      W_g[13,37] := -0.07636662;
      W_g[13,38] := -0.02541909;
      W_g[13,39] := -0.00815807;
      W_g[14,0] := 0.05384851;
      W_g[14,1] := -0.08540776;
      W_g[14,2] := -0.08017597;
      W_g[14,3] := -0.28711280;
      W_g[14,4] := -0.38180253;
      W_g[14,5] := -0.12807073;
      W_g[14,6] := -0.33112118;
      W_g[14,7] := -0.01536665;
      W_g[14,8] := 0.07860034;
      W_g[14,9] := 0.07597807;
      W_g[14,10] := 0.81271881;
      W_g[14,11] := 0.34440023;
      W_g[14,12] := -0.11264267;
      W_g[14,13] := 0.29767352;
      W_g[14,14] := -0.05823113;
      W_g[14,15] := -0.00107844;
      W_g[14,16] := -0.02762355;
      W_g[14,17] := -0.02232336;
      W_g[14,18] := 0.03123496;
      W_g[14,19] := -0.13857344;
      W_g[14,20] := 0.10911304;
      W_g[14,21] := -0.12785229;
      W_g[14,22] := -0.04815350;
      W_g[14,23] := -0.17390981;
      W_g[14,24] := 0.13923632;
      W_g[14,25] := 0.11850380;
      W_g[14,26] := -0.32757759;
      W_g[14,27] := -0.25137767;
      W_g[14,28] := 0.22421645;
      W_g[14,29] := -0.42832899;
      W_g[14,30] := 0.06481594;
      W_g[14,31] := -0.23915793;
      W_g[14,32] := -0.04046796;
      W_g[14,33] := -0.09582479;
      W_g[14,34] := -0.09370243;
      W_g[14,35] := 0.14524275;
      W_g[14,36] := -0.03895468;
      W_g[14,37] := 0.10286443;
      W_g[14,38] := 0.03800159;
      W_g[14,39] := 0.11008195;
      W_g[15,0] := 0.49670509;
      W_g[15,1] := 0.19451231;
      W_g[15,2] := -0.24881296;
      W_g[15,3] := 0.56299460;
      W_g[15,4] := -0.14983681;
      W_g[15,5] := -0.02904006;
      W_g[15,6] := 0.06259420;
      W_g[15,7] := 0.16642898;
      W_g[15,8] := -0.08521152;
      W_g[15,9] := -0.12409624;
      W_g[15,10] := 0.24281517;
      W_g[15,11] := -0.10940242;
      W_g[15,12] := 0.71269953;
      W_g[15,13] := -0.18780579;
      W_g[15,14] := 0.00091037;
      W_g[15,15] := -0.06534981;
      W_g[15,16] := 0.00326133;
      W_g[15,17] := -0.00118504;
      W_g[15,18] := -0.04420842;
      W_g[15,19] := -0.22520956;
      W_g[15,20] := -0.11959776;
      W_g[15,21] := -0.10079119;
      W_g[15,22] := -0.04329386;
      W_g[15,23] := -0.07395163;
      W_g[15,24] := -0.11715485;
      W_g[15,25] := -0.18832952;
      W_g[15,26] := -0.24700920;
      W_g[15,27] := -0.09096922;
      W_g[15,28] := 0.07692285;
      W_g[15,29] := 0.01714239;
      W_g[15,30] := -0.08180999;
      W_g[15,31] := -0.00006038;
      W_g[15,32] := 0.02792178;
      W_g[15,33] := 0.08978129;
      W_g[15,34] := -0.02846152;
      W_g[15,35] := 0.05397168;
      W_g[15,36] := 0.01382420;
      W_g[15,37] := 0.12623927;
      W_g[15,38] := 0.02842882;
      W_g[15,39] := -0.23873122;
      W_g[16,0] := 0.00714069;
      W_g[16,1] := 0.09252225;
      W_g[16,2] := -0.01911032;
      W_g[16,3] := 0.04820935;
      W_g[16,4] := 0.04210250;
      W_g[16,5] := 0.05442985;
      W_g[16,6] := 0.24199863;
      W_g[16,7] := -0.08810946;
      W_g[16,8] := 0.02272573;
      W_g[16,9] := -0.01153773;
      W_g[16,10] := -0.01938002;
      W_g[16,11] := 0.95534259;
      W_g[16,12] := 0.00685452;
      W_g[16,13] := -0.05267539;
      W_g[16,14] := -0.04784015;
      W_g[16,15] := 0.02123881;
      W_g[16,16] := 0.02990256;
      W_g[16,17] := 0.22012618;
      W_g[16,18] := -0.12446024;
      W_g[16,19] := 0.01318580;
      W_g[16,20] := 0.31736228;
      W_g[16,21] := 0.25552613;
      W_g[16,22] := 0.02996899;
      W_g[16,23] := 0.13324806;
      W_g[16,24] := 0.01029211;
      W_g[16,25] := -0.11731086;
      W_g[16,26] := 0.08171849;
      W_g[16,27] := -0.11919475;
      W_g[16,28] := 0.04512075;
      W_g[16,29] := 0.04511562;
      W_g[16,30] := 0.01768237;
      W_g[16,31] := -0.11807074;
      W_g[16,32] := 0.02917237;
      W_g[16,33] := 0.08451862;
      W_g[16,34] := 0.18420373;
      W_g[16,35] := 0.06097095;
      W_g[16,36] := 0.01656622;
      W_g[16,37] := -0.02950481;
      W_g[16,38] := 0.00875620;
      W_g[16,39] := -0.30139515;
      W_g[17,0] := 0.28211352;
      W_g[17,1] := -0.06947739;
      W_g[17,2] := -0.48255709;
      W_g[17,3] := -0.48009890;
      W_g[17,4] := 0.40037093;
      W_g[17,5] := -0.41533524;
      W_g[17,6] := 0.61539871;
      W_g[17,7] := -0.07803038;
      W_g[17,8] := 0.20740844;
      W_g[17,9] := 0.19454060;
      W_g[17,10] := 0.37828967;
      W_g[17,11] := 0.51134646;
      W_g[17,12] := 0.02942824;
      W_g[17,13] := -0.03419436;
      W_g[17,14] := -0.14622004;
      W_g[17,15] := 0.12808461;
      W_g[17,16] := -0.08771772;
      W_g[17,17] := -0.17915098;
      W_g[17,18] := -0.35652786;
      W_g[17,19] := -0.08436973;
      W_g[17,20] := -0.15241621;
      W_g[17,21] := -0.59241575;
      W_g[17,22] := -0.12622987;
      W_g[17,23] := -0.06875754;
      W_g[17,24] := -0.61650282;
      W_g[17,25] := -0.62400168;
      W_g[17,26] := 0.12978441;
      W_g[17,27] := 0.19093341;
      W_g[17,28] := -0.57437402;
      W_g[17,29] := -0.10343723;
      W_g[17,30] := -0.14047481;
      W_g[17,31] := 0.10861561;
      W_g[17,32] := -0.08338292;
      W_g[17,33] := -0.15795745;
      W_g[17,34] := -1.05674601;
      W_g[17,35] := 0.07798125;
      W_g[17,36] := -0.04106956;
      W_g[17,37] := -0.14353254;
      W_g[17,38] := -0.01768998;
      W_g[17,39] := 0.23552968;
      W_g[18,0] := -0.56118143;
      W_g[18,1] := 0.01680752;
      W_g[18,2] := 0.21060835;
      W_g[18,3] := 0.22311090;
      W_g[18,4] := -0.35391527;
      W_g[18,5] := -0.00398842;
      W_g[18,6] := 0.44133097;
      W_g[18,7] := -0.20236395;
      W_g[18,8] := 0.27059153;
      W_g[18,9] := -0.26535335;
      W_g[18,10] := -0.00161409;
      W_g[18,11] := -0.42498562;
      W_g[18,12] := 0.18595842;
      W_g[18,13] := 0.03403796;
      W_g[18,14] := -0.19036941;
      W_g[18,15] := 0.00153053;
      W_g[18,16] := -0.13208415;
      W_g[18,17] := -0.00688618;
      W_g[18,18] := 0.04695740;
      W_g[18,19] := 0.52580279;
      W_g[18,20] := 0.33302781;
      W_g[18,21] := -0.03863472;
      W_g[18,22] := -0.04098545;
      W_g[18,23] := 0.05270698;
      W_g[18,24] := -0.87936115;
      W_g[18,25] := -0.79176319;
      W_g[18,26] := -0.37981445;
      W_g[18,27] := -0.39054155;
      W_g[18,28] := 0.40099201;
      W_g[18,29] := -0.21964216;
      W_g[18,30] := -0.06956752;
      W_g[18,31] := 1.08965826;
      W_g[18,32] := -0.24863915;
      W_g[18,33] := 0.04124767;
      W_g[18,34] := -0.14617871;
      W_g[18,35] := -0.54955792;
      W_g[18,36] := 0.22360204;
      W_g[18,37] := -0.51476938;
      W_g[18,38] := -0.00649375;
      W_g[18,39] := 0.23745580;
      W_g[19,0] := 0.04427215;
      W_g[19,1] := 0.13209015;
      W_g[19,2] := -0.12966105;
      W_g[19,3] := 0.13671713;
      W_g[19,4] := 0.01762369;
      W_g[19,5] := 0.09627694;
      W_g[19,6] := -0.13640797;
      W_g[19,7] := 0.02292525;
      W_g[19,8] := 0.06818993;
      W_g[19,9] := -0.01616117;
      W_g[19,10] := -0.27115190;
      W_g[19,11] := -0.17511748;
      W_g[19,12] := 0.20083658;
      W_g[19,13] := 0.12117302;
      W_g[19,14] := -0.40477425;
      W_g[19,15] := 0.00942509;
      W_g[19,16] := -0.00977145;
      W_g[19,17] := -0.00656325;
      W_g[19,18] := -0.02440832;
      W_g[19,19] := -0.10208004;
      W_g[19,20] := 0.05442004;
      W_g[19,21] := -0.28210428;
      W_g[19,22] := -0.02802154;
      W_g[19,23] := -0.16558743;
      W_g[19,24] := 0.24839798;
      W_g[19,25] := 0.68076271;
      W_g[19,26] := -0.15649894;
      W_g[19,27] := 0.02872765;
      W_g[19,28] := -0.14855081;
      W_g[19,29] := -0.04783039;
      W_g[19,30] := -0.04433315;
      W_g[19,31] := -0.00463518;
      W_g[19,32] := -0.04792630;
      W_g[19,33] := -0.18936750;
      W_g[19,34] := -0.28109401;
      W_g[19,35] := 0.12269117;
      W_g[19,36] := -0.02590044;
      W_g[19,37] := 0.13191973;
      W_g[19,38] := -0.08906776;
      W_g[19,39] := -0.30020091;
      W_g[20,0] := -0.20718005;
      W_g[20,1] := -0.84034145;
      W_g[20,2] := 0.02167286;
      W_g[20,3] := 0.22337365;
      W_g[20,4] := -0.22535181;
      W_g[20,5] := 0.00862414;
      W_g[20,6] := -0.07585888;
      W_g[20,7] := 0.20224823;
      W_g[20,8] := 0.33609936;
      W_g[20,9] := 0.24086921;
      W_g[20,10] := -0.34230143;
      W_g[20,11] := 0.23271726;
      W_g[20,12] := -0.54696190;
      W_g[20,13] := 0.07557353;
      W_g[20,14] := -0.00750887;
      W_g[20,15] := -0.07179558;
      W_g[20,16] := 0.11929045;
      W_g[20,17] := 0.01187360;
      W_g[20,18] := 0.01727761;
      W_g[20,19] := -0.10120918;
      W_g[20,20] := -0.35278231;
      W_g[20,21] := -0.09405834;
      W_g[20,22] := 0.04689666;
      W_g[20,23] := -0.10715894;
      W_g[20,24] := -0.07375087;
      W_g[20,25] := -0.14543816;
      W_g[20,26] := -0.23896208;
      W_g[20,27] := -0.43519315;
      W_g[20,28] := -0.25828305;
      W_g[20,29] := -0.05447736;
      W_g[20,30] := 0.05642707;
      W_g[20,31] := 0.18183576;
      W_g[20,32] := 0.08492490;
      W_g[20,33] := 0.19067700;
      W_g[20,34] := -0.11871803;
      W_g[20,35] := -0.03175204;
      W_g[20,36] := -0.04638923;
      W_g[20,37] := -0.03955484;
      W_g[20,38] := 0.18262649;
      W_g[20,39] := -0.00053967;
      W_g[21,0] := -0.00852127;
      W_g[21,1] := 0.16749823;
      W_g[21,2] := -0.15172872;
      W_g[21,3] := -0.20800257;
      W_g[21,4] := 0.15032937;
      W_g[21,5] := 0.06710505;
      W_g[21,6] := -0.26149949;
      W_g[21,7] := 0.03740874;
      W_g[21,8] := 0.13018388;
      W_g[21,9] := 0.18329854;
      W_g[21,10] := -0.03891287;
      W_g[21,11] := 0.05188271;
      W_g[21,12] := 0.47803098;
      W_g[21,13] := 0.06662370;
      W_g[21,14] := -0.00612103;
      W_g[21,15] := -0.13870122;
      W_g[21,16] := -0.10494442;
      W_g[21,17] := -0.00346555;
      W_g[21,18] := -0.04227602;
      W_g[21,19] := -0.33476129;
      W_g[21,20] := 0.34089175;
      W_g[21,21] := 0.45425063;
      W_g[21,22] := 0.16435136;
      W_g[21,23] := 0.04143468;
      W_g[21,24] := 0.16786721;
      W_g[21,25] := 0.11948983;
      W_g[21,26] := 0.05792047;
      W_g[21,27] := -0.12976640;
      W_g[21,28] := -0.13790442;
      W_g[21,29] := 0.24387960;
      W_g[21,30] := 0.16521277;
      W_g[21,31] := 0.16834626;
      W_g[21,32] := -0.10805231;
      W_g[21,33] := -0.07898282;
      W_g[21,34] := 0.28881353;
      W_g[21,35] := -0.11385613;
      W_g[21,36] := -0.66726488;
      W_g[21,37] := -0.28654984;
      W_g[21,38] := 0.35271052;
      W_g[21,39] := 0.00955431;
      W_g[22,0] := 0.29109696;
      W_g[22,1] := 0.01384218;
      W_g[22,2] := -0.37709463;
      W_g[22,3] := 0.14574254;
      W_g[22,4] := -0.07661973;
      W_g[22,5] := 0.12081382;
      W_g[22,6] := -0.39220569;
      W_g[22,7] := -0.00977318;
      W_g[22,8] := 0.02812388;
      W_g[22,9] := -0.07591717;
      W_g[22,10] := -0.08413436;
      W_g[22,11] := 0.17591499;
      W_g[22,12] := -0.33312052;
      W_g[22,13] := -0.12893844;
      W_g[22,14] := 0.12280960;
      W_g[22,15] := 0.33149692;
      W_g[22,16] := -0.12770943;
      W_g[22,17] := 0.11019890;
      W_g[22,18] := -0.02004679;
      W_g[22,19] := -0.09840271;
      W_g[22,20] := -0.03289499;
      W_g[22,21] := -0.03317460;
      W_g[22,22] := 0.05239879;
      W_g[22,23] := 0.39912307;
      W_g[22,24] := 0.28896907;
      W_g[22,25] := -0.06105658;
      W_g[22,26] := -0.21285506;
      W_g[22,27] := -0.03863349;
      W_g[22,28] := 0.16256362;
      W_g[22,29] := 0.14152323;
      W_g[22,30] := 0.05700575;
      W_g[22,31] := 0.37323594;
      W_g[22,32] := -0.00197801;
      W_g[22,33] := 0.01016807;
      W_g[22,34] := -0.05393393;
      W_g[22,35] := -0.03373878;
      W_g[22,36] := 0.00123443;
      W_g[22,37] := -0.10641941;
      W_g[22,38] := -0.03629038;
      W_g[22,39] := -0.09397990;
      W_g[23,0] := -0.09347695;
      W_g[23,1] := -0.22505829;
      W_g[23,2] := 0.01111710;
      W_g[23,3] := -0.13649231;
      W_g[23,4] := -0.30517000;
      W_g[23,5] := 0.83911264;
      W_g[23,6] := -0.75282311;
      W_g[23,7] := -0.66691148;
      W_g[23,8] := 0.15447931;
      W_g[23,9] := -0.55708647;
      W_g[23,10] := 0.25686628;
      W_g[23,11] := 0.12212675;
      W_g[23,12] := 0.16343321;
      W_g[23,13] := -0.31660068;
      W_g[23,14] := 0.02282131;
      W_g[23,15] := -0.05205119;
      W_g[23,16] := -0.05839873;
      W_g[23,17] := -0.09075660;
      W_g[23,18] := -0.23147778;
      W_g[23,19] := 0.07263616;
      W_g[23,20] := -0.51794368;
      W_g[23,21] := -0.27791360;
      W_g[23,22] := -0.07805633;
      W_g[23,23] := -0.41355452;
      W_g[23,24] := -0.21751262;
      W_g[23,25] := -0.05684796;
      W_g[23,26] := 0.30686048;
      W_g[23,27] := -0.14003992;
      W_g[23,28] := -0.38135511;
      W_g[23,29] := 0.13330600;
      W_g[23,30] := -0.06790695;
      W_g[23,31] := -0.07987443;
      W_g[23,32] := 0.06365003;
      W_g[23,33] := 0.22799088;
      W_g[23,34] := 0.13270302;
      W_g[23,35] := -0.00725970;
      W_g[23,36] := 0.16376778;
      W_g[23,37] := -0.02287991;
      W_g[23,38] := 0.08711061;
      W_g[23,39] := 0.01950686;
      W_g[24,0] := 0.46194655;
      W_g[24,1] := 0.27763960;
      W_g[24,2] := -0.12869456;
      W_g[24,3] := 0.13782990;
      W_g[24,4] := -1.03041399;
      W_g[24,5] := 0.00441816;
      W_g[24,6] := 0.44230226;
      W_g[24,7] := 0.18489341;
      W_g[24,8] := -0.30371043;
      W_g[24,9] := 0.03693367;
      W_g[24,10] := -0.01524317;
      W_g[24,11] := -0.24215870;
      W_g[24,12] := 0.35080424;
      W_g[24,13] := 0.07174128;
      W_g[24,14] := 0.00412538;
      W_g[24,15] := 0.02062515;
      W_g[24,16] := 0.01971583;
      W_g[24,17] := 0.00580471;
      W_g[24,18] := -0.04475251;
      W_g[24,19] := -0.08863095;
      W_g[24,20] := 0.06659620;
      W_g[24,21] := -0.19372395;
      W_g[24,22] := 0.04916465;
      W_g[24,23] := 0.11263776;
      W_g[24,24] := 0.45533353;
      W_g[24,25] := 0.28435835;
      W_g[24,26] := 0.23480317;
      W_g[24,27] := -0.41078931;
      W_g[24,28] := -0.25990930;
      W_g[24,29] := 0.04082377;
      W_g[24,30] := 0.05907518;
      W_g[24,31] := 0.00033808;
      W_g[24,32] := -0.03658906;
      W_g[24,33] := -0.08924066;
      W_g[24,34] := -0.02038150;
      W_g[24,35] := 0.01517213;
      W_g[24,36] := -0.29084125;
      W_g[24,37] := -0.03483975;
      W_g[24,38] := -0.33877048;
      W_g[24,39] := 0.01846378;
      W_g[25,0] := -0.01319884;
      W_g[25,1] := 0.17892542;
      W_g[25,2] := 0.00354903;
      W_g[25,3] := -0.01092031;
      W_g[25,4] := 0.04581180;
      W_g[25,5] := -0.04252854;
      W_g[25,6] := -0.05655812;
      W_g[25,7] := 0.07682356;
      W_g[25,8] := -0.01679150;
      W_g[25,9] := 0.05484685;
      W_g[25,10] := -0.09173104;
      W_g[25,11] := -0.12738757;
      W_g[25,12] := -0.10293069;
      W_g[25,13] := -0.00530847;
      W_g[25,14] := -0.08904938;
      W_g[25,15] := 0.36966512;
      W_g[25,16] := -0.00969987;
      W_g[25,17] := -0.28969538;
      W_g[25,18] := -0.02469883;
      W_g[25,19] := -0.08574332;
      W_g[25,20] := 0.10813141;
      W_g[25,21] := 0.08889347;
      W_g[25,22] := -0.06467538;
      W_g[25,23] := 0.04102366;
      W_g[25,24] := -0.24661052;
      W_g[25,25] := -0.24702097;
      W_g[25,26] := -0.08217103;
      W_g[25,27] := -0.05707087;
      W_g[25,28] := -0.01940200;
      W_g[25,29] := -0.00729063;
      W_g[25,30] := -0.06900500;
      W_g[25,31] := -0.19478676;
      W_g[25,32] := 0.08665588;
      W_g[25,33] := 0.17711434;
      W_g[25,34] := 0.35117847;
      W_g[25,35] := 0.00400291;
      W_g[25,36] := 0.02780187;
      W_g[25,37] := -0.02507502;
      W_g[25,38] := 0.01814217;
      W_g[25,39] := 0.01270028;
      W_g[26,0] := -0.10013371;
      W_g[26,1] := -0.11928739;
      W_g[26,2] := 0.03542966;
      W_g[26,3] := -0.09299100;
      W_g[26,4] := 0.22154348;
      W_g[26,5] := 0.04870279;
      W_g[26,6] := -0.01336484;
      W_g[26,7] := -0.05781888;
      W_g[26,8] := 0.00065369;
      W_g[26,9] := -0.01473211;
      W_g[26,10] := -0.01971318;
      W_g[26,11] := 0.02451181;
      W_g[26,12] := 0.14100704;
      W_g[26,13] := 0.20081082;
      W_g[26,14] := -0.00175938;
      W_g[26,15] := -0.13420245;
      W_g[26,16] := 0.01900839;
      W_g[26,17] := -0.02341681;
      W_g[26,18] := -0.94101948;
      W_g[26,19] := -0.02586854;
      W_g[26,20] := -0.30304915;
      W_g[26,21] := 0.06037450;
      W_g[26,22] := -0.02225667;
      W_g[26,23] := 0.34992269;
      W_g[26,24] := -0.15178578;
      W_g[26,25] := -0.21104257;
      W_g[26,26] := -0.25511426;
      W_g[26,27] := -0.03610617;
      W_g[26,28] := -0.13982570;
      W_g[26,29] := -0.07677662;
      W_g[26,30] := -0.02899644;
      W_g[26,31] := 0.02322534;
      W_g[26,32] := -0.01148466;
      W_g[26,33] := 0.01643471;
      W_g[26,34] := -0.05193237;
      W_g[26,35] := -0.01343275;
      W_g[26,36] := 0.01284295;
      W_g[26,37] := 0.01176736;
      W_g[26,38] := 0.00468252;
      W_g[26,39] := -0.20358260;
      W_g[27,0] := 0.01242287;
      W_g[27,1] := -0.01930982;
      W_g[27,2] := -0.24737412;
      W_g[27,3] := -0.13776387;
      W_g[27,4] := 0.19126348;
      W_g[27,5] := 0.00086061;
      W_g[27,6] := -0.16852112;
      W_g[27,7] := -0.08134060;
      W_g[27,8] := 0.29883468;
      W_g[27,9] := 0.09754812;
      W_g[27,10] := 0.09034698;
      W_g[27,11] := -0.06812658;
      W_g[27,12] := -0.14695419;
      W_g[27,13] := -0.05109974;
      W_g[27,14] := -0.01788860;
      W_g[27,15] := -0.15783192;
      W_g[27,16] := 0.19530444;
      W_g[27,17] := -0.16005373;
      W_g[27,18] := 0.26013258;
      W_g[27,19] := 0.26764771;
      W_g[27,20] := -0.12696983;
      W_g[27,21] := 0.31249490;
      W_g[27,22] := 0.09300645;
      W_g[27,23] := 0.03466551;
      W_g[27,24] := 0.23168693;
      W_g[27,25] := 0.18956751;
      W_g[27,26] := -0.04334988;
      W_g[27,27] := -0.18214862;
      W_g[27,28] := -0.04629618;
      W_g[27,29] := 0.09379144;
      W_g[27,30] := 0.07671305;
      W_g[27,31] := -0.01221954;
      W_g[27,32] := -0.02424719;
      W_g[27,33] := 0.07423434;
      W_g[27,34] := 0.18019708;
      W_g[27,35] := -0.04701952;
      W_g[27,36] := -0.08283819;
      W_g[27,37] := -0.09333491;
      W_g[27,38] := -0.48927879;
      W_g[27,39] := -0.00745687;
      W_g[28,0] := 0.13821959;
      W_g[28,1] := 0.07419970;
      W_g[28,2] := -0.28731343;
      W_g[28,3] := 0.52230597;
      W_g[28,4] := 0.13792820;
      W_g[28,5] := -0.04003582;
      W_g[28,6] := 0.12009837;
      W_g[28,7] := -0.22427090;
      W_g[28,8] := 0.10034105;
      W_g[28,9] := -0.43725863;
      W_g[28,10] := 0.10780185;
      W_g[28,11] := -0.03007025;
      W_g[28,12] := -0.09082274;
      W_g[28,13] := 0.21732096;
      W_g[28,14] := -0.03366475;
      W_g[28,15] := 0.12757394;
      W_g[28,16] := 0.40819040;
      W_g[28,17] := 0.08709385;
      W_g[28,18] := -0.01960146;
      W_g[28,19] := -0.01771599;
      W_g[28,20] := 0.02389354;
      W_g[28,21] := 0.04893105;
      W_g[28,22] := 0.01708278;
      W_g[28,23] := 0.05532730;
      W_g[28,24] := -0.42513239;
      W_g[28,25] := -0.53693467;
      W_g[28,26] := 0.09680068;
      W_g[28,27] := 0.11012019;
      W_g[28,28] := -0.10853667;
      W_g[28,29] := -0.10696560;
      W_g[28,30] := -0.01152095;
      W_g[28,31] := 0.08765919;
      W_g[28,32] := -0.04124034;
      W_g[28,33] := 0.00073121;
      W_g[28,34] := -0.07680846;
      W_g[28,35] := -0.09583755;
      W_g[28,36] := -0.02250235;
      W_g[28,37] := -0.10466012;
      W_g[28,38] := 0.02804276;
      W_g[28,39] := 0.05010757;
      W_g[29,0] := -0.13576494;
      W_g[29,1] := -0.04743524;
      W_g[29,2] := 0.01165335;
      W_g[29,3] := -0.06858198;
      W_g[29,4] := 0.11698179;
      W_g[29,5] := 0.15293106;
      W_g[29,6] := -0.08868138;
      W_g[29,7] := 0.00604072;
      W_g[29,8] := 0.10700601;
      W_g[29,9] := 0.08990686;
      W_g[29,10] := -0.17016383;
      W_g[29,11] := -0.09298281;
      W_g[29,12] := 0.23396063;
      W_g[29,13] := -0.43684760;
      W_g[29,14] := -0.02256006;
      W_g[29,15] := 0.02156748;
      W_g[29,16] := -0.04530424;
      W_g[29,17] := 0.02112582;
      W_g[29,18] := 0.43311554;
      W_g[29,19] := 0.28956264;
      W_g[29,20] := -0.45648861;
      W_g[29,21] := -0.47465628;
      W_g[29,22] := -0.15953651;
      W_g[29,23] := 0.62224460;
      W_g[29,24] := -0.36037850;
      W_g[29,25] := -0.32347810;
      W_g[29,26] := -0.10036322;
      W_g[29,27] := 0.23475674;
      W_g[29,28] := -0.38871291;
      W_g[29,29] := -0.37588716;
      W_g[29,30] := -0.19999301;
      W_g[29,31] := -0.07129297;
      W_g[29,32] := 0.00924866;
      W_g[29,33] := -0.00100953;
      W_g[29,34] := -0.03974389;
      W_g[29,35] := 0.19243315;
      W_g[29,36] := -0.05763126;
      W_g[29,37] := 0.14980933;
      W_g[29,38] := 0.09773512;
      W_g[29,39] := 0.28358760;
      W_g[30,0] := 0.02073097;
      W_g[30,1] := -0.05142897;
      W_g[30,2] := 0.05679109;
      W_g[30,3] := -0.29680440;
      W_g[30,4] := -0.09398746;
      W_g[30,5] := 0.00418108;
      W_g[30,6] := -0.12116858;
      W_g[30,7] := 0.13785014;
      W_g[30,8] := -0.07182530;
      W_g[30,9] := 0.28989494;
      W_g[30,10] := -0.02703100;
      W_g[30,11] := -0.04196686;
      W_g[30,12] := 0.23686379;
      W_g[30,13] := -0.11817347;
      W_g[30,14] := -0.00608444;
      W_g[30,15] := 0.27866739;
      W_g[30,16] := 0.31624600;
      W_g[30,17] := -0.04371030;
      W_g[30,18] := -0.09872175;
      W_g[30,19] := 0.17183733;
      W_g[30,20] := -0.10328431;
      W_g[30,21] := 0.02654029;
      W_g[30,22] := 0.04664133;
      W_g[30,23] := -0.02138521;
      W_g[30,24] := 0.42544174;
      W_g[30,25] := -0.03961691;
      W_g[30,26] := 0.11087703;
      W_g[30,27] := 0.09755427;
      W_g[30,28] := 0.11475538;
      W_g[30,29] := 0.06603787;
      W_g[30,30] := 0.05809331;
      W_g[30,31] := 0.13511968;
      W_g[30,32] := -0.00735715;
      W_g[30,33] := -0.00152808;
      W_g[30,34] := -0.12982640;
      W_g[30,35] := 0.00118882;
      W_g[30,36] := 0.01855830;
      W_g[30,37] := -0.05438844;
      W_g[30,38] := 0.05046400;
      W_g[30,39] := -0.03010074;
      W_g[31,0] := 0.08256169;
      W_g[31,1] := -0.51133311;
      W_g[31,2] := 0.11336197;
      W_g[31,3] := -0.15730928;
      W_g[31,4] := 0.15212694;
      W_g[31,5] := 0.05411269;
      W_g[31,6] := -0.07535803;
      W_g[31,7] := 0.03512096;
      W_g[31,8] := -0.05313810;
      W_g[31,9] := 0.10365095;
      W_g[31,10] := -0.00368842;
      W_g[31,11] := -0.12890872;
      W_g[31,12] := 0.47981134;
      W_g[31,13] := 0.03815160;
      W_g[31,14] := -0.01872904;
      W_g[31,15] := 0.17062889;
      W_g[31,16] := -0.12828785;
      W_g[31,17] := 0.06558654;
      W_g[31,18] := -0.06244295;
      W_g[31,19] := -0.53075397;
      W_g[31,20] := 0.15929437;
      W_g[31,21] := 0.00589449;
      W_g[31,22] := -0.03731958;
      W_g[31,23] := 0.05464490;
      W_g[31,24] := -0.19547676;
      W_g[31,25] := 0.11578897;
      W_g[31,26] := 0.27690557;
      W_g[31,27] := 0.26996168;
      W_g[31,28] := 0.03783383;
      W_g[31,29] := -0.16668507;
      W_g[31,30] := -0.05871727;
      W_g[31,31] := 0.11560699;
      W_g[31,32] := -0.10597849;
      W_g[31,33] := -0.03747635;
      W_g[31,34] := -0.06264409;
      W_g[31,35] := -0.18381201;
      W_g[31,36] := 0.07526756;
      W_g[31,37] := -0.11970815;
      W_g[31,38] := -0.33985323;
      W_g[31,39] := 0.02983656;
      W_o[0,0] := 0.13366428;
      W_o[0,1] := 0.11036980;
      W_o[0,2] := -0.16846675;
      W_o[0,3] := -0.21495235;
      W_o[0,4] := 0.07811608;
      W_o[0,5] := -0.13181226;
      W_o[0,6] := -0.32309711;
      W_o[0,7] := -0.05775660;
      W_o[0,8] := 0.07714970;
      W_o[0,9] := 0.69965583;
      W_o[0,10] := 0.03330577;
      W_o[0,11] := 0.07725812;
      W_o[0,12] := 0.25551820;
      W_o[0,13] := 0.38036522;
      W_o[0,14] := -0.01993838;
      W_o[0,15] := -0.05171372;
      W_o[0,16] := 0.00189644;
      W_o[0,17] := -0.32097366;
      W_o[0,18] := -0.05273939;
      W_o[0,19] := 0.04321737;
      W_o[0,20] := -0.23801146;
      W_o[0,21] := 0.29699677;
      W_o[0,22] := -0.16276316;
      W_o[0,23] := -0.23706993;
      W_o[0,24] := 0.17703076;
      W_o[0,25] := 0.36713782;
      W_o[0,26] := -0.12915254;
      W_o[0,27] := -0.07524700;
      W_o[0,28] := -0.09860305;
      W_o[0,29] := 0.12421684;
      W_o[0,30] := -0.39039981;
      W_o[0,31] := -0.01002511;
      W_o[0,32] := -0.46100792;
      W_o[0,33] := 0.17252544;
      W_o[0,34] := 0.15642625;
      W_o[0,35] := -0.27402765;
      W_o[0,36] := -0.07788435;
      W_o[0,37] := -0.09713101;
      W_o[0,38] := -0.05069508;
      W_o[0,39] := -0.24549620;
      W_o[1,0] := 0.49653649;
      W_o[1,1] := -0.05346184;
      W_o[1,2] := -0.01993282;
      W_o[1,3] := -0.13199322;
      W_o[1,4] := 0.03771848;
      W_o[1,5] := 0.14309798;
      W_o[1,6] := 0.04961836;
      W_o[1,7] := 0.27153552;
      W_o[1,8] := 0.60058177;
      W_o[1,9] := -0.62969673;
      W_o[1,10] := 0.21819758;
      W_o[1,11] := -0.10272143;
      W_o[1,12] := 0.11986823;
      W_o[1,13] := -0.24452005;
      W_o[1,14] := -0.06335072;
      W_o[1,15] := -0.16848719;
      W_o[1,16] := -0.21195354;
      W_o[1,17] := 0.02550812;
      W_o[1,18] := -0.14588526;
      W_o[1,19] := -0.51397264;
      W_o[1,20] := -0.21644965;
      W_o[1,21] := -0.53661948;
      W_o[1,22] := -0.02092957;
      W_o[1,23] := 0.01972848;
      W_o[1,24] := -0.55939800;
      W_o[1,25] := -0.49083781;
      W_o[1,26] := -0.14633974;
      W_o[1,27] := 0.42070836;
      W_o[1,28] := -0.21612938;
      W_o[1,29] := -0.03745779;
      W_o[1,30] := 0.06127948;
      W_o[1,31] := 0.35676870;
      W_o[1,32] := -0.08789702;
      W_o[1,33] := 0.11810053;
      W_o[1,34] := -0.01725286;
      W_o[1,35] := -0.06969324;
      W_o[1,36] := -0.01398361;
      W_o[1,37] := -0.15410708;
      W_o[1,38] := -0.08071988;
      W_o[1,39] := -0.25934911;
      W_o[2,0] := 0.13397244;
      W_o[2,1] := -0.67044854;
      W_o[2,2] := -0.32567781;
      W_o[2,3] := -0.75043666;
      W_o[2,4] := -0.32291642;
      W_o[2,5] := 0.54297352;
      W_o[2,6] := 1.01406825;
      W_o[2,7] := -0.63293743;
      W_o[2,8] := -0.24675053;
      W_o[2,9] := -0.54400074;
      W_o[2,10] := -0.70754099;
      W_o[2,11] := -0.16770625;
      W_o[2,12] := -0.13771380;
      W_o[2,13] := -0.93835974;
      W_o[2,14] := 0.07016375;
      W_o[2,15] := -0.14486392;
      W_o[2,16] := 0.26753914;
      W_o[2,17] := -0.44003579;
      W_o[2,18] := -0.19662693;
      W_o[2,19] := 0.14748774;
      W_o[2,20] := 0.04340832;
      W_o[2,21] := 0.91405821;
      W_o[2,22] := 0.23963371;
      W_o[2,23] := -0.42069820;
      W_o[2,24] := 1.35907292;
      W_o[2,25] := 0.74127895;
      W_o[2,26] := -0.60126311;
      W_o[2,27] := 1.04573679;
      W_o[2,28] := 0.35571697;
      W_o[2,29] := 0.19770171;
      W_o[2,30] := 0.19496830;
      W_o[2,31] := -0.06545950;
      W_o[2,32] := -0.07142299;
      W_o[2,33] := -0.23412317;
      W_o[2,34] := 0.13213682;
      W_o[2,35] := 0.09960951;
      W_o[2,36] := -0.82927501;
      W_o[2,37] := -0.00553483;
      W_o[2,38] := 0.72544241;
      W_o[2,39] := 0.20440662;
      W_o[3,0] := -0.29025504;
      W_o[3,1] := 0.21485890;
      W_o[3,2] := 0.12162556;
      W_o[3,3] := -0.45000923;
      W_o[3,4] := 0.00440878;
      W_o[3,5] := -0.07761150;
      W_o[3,6] := 0.27128229;
      W_o[3,7] := 0.20583764;
      W_o[3,8] := 0.36606720;
      W_o[3,9] := 0.31630817;
      W_o[3,10] := 0.16728929;
      W_o[3,11] := 0.21024089;
      W_o[3,12] := -0.30256730;
      W_o[3,13] := -0.07960982;
      W_o[3,14] := 0.26832253;
      W_o[3,15] := 0.38332802;
      W_o[3,16] := 0.01548071;
      W_o[3,17] := 0.27411333;
      W_o[3,18] := -0.07721005;
      W_o[3,19] := -0.15753639;
      W_o[3,20] := -0.12283424;
      W_o[3,21] := -0.09994975;
      W_o[3,22] := -0.25781667;
      W_o[3,23] := -0.30848202;
      W_o[3,24] := 0.08977263;
      W_o[3,25] := -0.00644524;
      W_o[3,26] := 0.31200859;
      W_o[3,27] := -0.01467965;
      W_o[3,28] := -0.12804723;
      W_o[3,29] := -0.06573117;
      W_o[3,30] := -0.39431822;
      W_o[3,31] := -0.44901580;
      W_o[3,32] := -0.13384379;
      W_o[3,33] := -0.10575464;
      W_o[3,34] := 0.01442572;
      W_o[3,35] := -0.11673454;
      W_o[3,36] := -0.14822102;
      W_o[3,37] := -0.02524356;
      W_o[3,38] := -0.03832110;
      W_o[3,39] := 0.94678485;
      W_o[4,0] := -0.89165902;
      W_o[4,1] := -0.07221486;
      W_o[4,2] := 0.45090771;
      W_o[4,3] := 0.40743887;
      W_o[4,4] := -0.00022854;
      W_o[4,5] := -0.22787750;
      W_o[4,6] := 0.56126112;
      W_o[4,7] := -0.65236539;
      W_o[4,8] := 0.31672934;
      W_o[4,9] := -0.60582823;
      W_o[4,10] := 0.85605830;
      W_o[4,11] := -0.86477047;
      W_o[4,12] := 0.63425988;
      W_o[4,13] := -0.08753718;
      W_o[4,14] := 0.07426148;
      W_o[4,15] := 0.43497530;
      W_o[4,16] := 0.02985676;
      W_o[4,17] := -0.01102423;
      W_o[4,18] := 0.00179447;
      W_o[4,19] := -0.39584765;
      W_o[4,20] := 0.37266934;
      W_o[4,21] := 0.29497612;
      W_o[4,22] := 0.37403074;
      W_o[4,23] := 0.22710080;
      W_o[4,24] := -1.35028052;
      W_o[4,25] := -0.25135967;
      W_o[4,26] := -0.09566695;
      W_o[4,27] := -0.22512139;
      W_o[4,28] := -0.06946037;
      W_o[4,29] := 0.32004294;
      W_o[4,30] := 0.36742997;
      W_o[4,31] := -0.14018387;
      W_o[4,32] := 0.11306093;
      W_o[4,33] := -0.10145790;
      W_o[4,34] := -0.10018518;
      W_o[4,35] := 0.20776151;
      W_o[4,36] := 0.04030388;
      W_o[4,37] := 0.23607983;
      W_o[4,38] := -0.00676852;
      W_o[4,39] := -0.01103176;
      W_o[5,0] := -0.13071172;
      W_o[5,1] := 0.17688261;
      W_o[5,2] := 0.09693976;
      W_o[5,3] := -0.24016836;
      W_o[5,4] := -0.17199296;
      W_o[5,5] := -0.06652235;
      W_o[5,6] := -0.37081853;
      W_o[5,7] := 0.06624742;
      W_o[5,8] := -0.20348907;
      W_o[5,9] := -0.21328829;
      W_o[5,10] := 0.18360765;
      W_o[5,11] := 0.27653855;
      W_o[5,12] := -0.57717568;
      W_o[5,13] := -0.11226647;
      W_o[5,14] := -0.08564992;
      W_o[5,15] := 0.21546762;
      W_o[5,16] := -0.33327058;
      W_o[5,17] := 0.02841459;
      W_o[5,18] := -0.26086703;
      W_o[5,19] := 0.29187077;
      W_o[5,20] := -0.36725804;
      W_o[5,21] := -0.09546806;
      W_o[5,22] := 0.45851558;
      W_o[5,23] := 0.07615964;
      W_o[5,24] := 1.94119501;
      W_o[5,25] := 1.68010128;
      W_o[5,26] := -0.03859005;
      W_o[5,27] := 0.21847658;
      W_o[5,28] := 0.21739782;
      W_o[5,29] := -0.10321381;
      W_o[5,30] := 0.33334309;
      W_o[5,31] := 0.09397009;
      W_o[5,32] := -0.12362885;
      W_o[5,33] := -0.02805139;
      W_o[5,34] := 0.22041477;
      W_o[5,35] := -0.33244985;
      W_o[5,36] := 0.18436120;
      W_o[5,37] := -0.52219701;
      W_o[5,38] := -0.11966625;
      W_o[5,39] := 0.01321488;
      W_o[6,0] := 0.25687075;
      W_o[6,1] := -0.82650340;
      W_o[6,2] := 0.32687336;
      W_o[6,3] := 0.02528367;
      W_o[6,4] := 0.15329729;
      W_o[6,5] := 0.29570559;
      W_o[6,6] := 0.89035386;
      W_o[6,7] := 0.05928367;
      W_o[6,8] := -0.37806994;
      W_o[6,9] := 0.04021226;
      W_o[6,10] := -0.35702997;
      W_o[6,11] := 0.21551481;
      W_o[6,12] := -0.07286788;
      W_o[6,13] := 0.37769529;
      W_o[6,14] := 0.00736793;
      W_o[6,15] := -0.05791439;
      W_o[6,16] := 0.23656519;
      W_o[6,17] := -0.04539794;
      W_o[6,18] := -0.00322705;
      W_o[6,19] := 0.23821436;
      W_o[6,20] := -1.42132485;
      W_o[6,21] := 0.48428133;
      W_o[6,22] := -0.18088701;
      W_o[6,23] := -0.22187343;
      W_o[6,24] := 1.33472562;
      W_o[6,25] := 0.99553061;
      W_o[6,26] := 0.20602396;
      W_o[6,27] := -0.03664935;
      W_o[6,28] := 0.17536840;
      W_o[6,29] := -0.02604117;
      W_o[6,30] := -0.18590604;
      W_o[6,31] := 0.00481638;
      W_o[6,32] := -0.31825411;
      W_o[6,33] := -0.24851917;
      W_o[6,34] := 0.63873190;
      W_o[6,35] := -0.29667321;
      W_o[6,36] := -0.02184569;
      W_o[6,37] := -0.29451790;
      W_o[6,38] := 0.29764518;
      W_o[6,39] := 0.21402869;
      W_o[7,0] := -1.12601244;
      W_o[7,1] := -0.86021799;
      W_o[7,2] := -1.00755525;
      W_o[7,3] := -0.12928128;
      W_o[7,4] := -0.41589841;
      W_o[7,5] := 0.27687931;
      W_o[7,6] := 0.24910082;
      W_o[7,7] := -0.15456890;
      W_o[7,8] := -1.40733433;
      W_o[7,9] := -0.16872104;
      W_o[7,10] := 0.02657967;
      W_o[7,11] := 0.15706138;
      W_o[7,12] := 0.48483267;
      W_o[7,13] := 0.17854783;
      W_o[7,14] := 0.01057731;
      W_o[7,15] := -0.06248428;
      W_o[7,16] := 0.01161261;
      W_o[7,17] := -0.04555431;
      W_o[7,18] := 0.78910136;
      W_o[7,19] := 0.23410527;
      W_o[7,20] := 0.23320967;
      W_o[7,21] := 0.44676164;
      W_o[7,22] := -0.00038366;
      W_o[7,23] := 0.21317144;
      W_o[7,24] := -0.20823158;
      W_o[7,25] := -0.08117293;
      W_o[7,26] := 0.15186004;
      W_o[7,27] := 0.05216801;
      W_o[7,28] := 0.74951005;
      W_o[7,29] := 0.27860886;
      W_o[7,30] := -0.01225667;
      W_o[7,31] := -0.13738722;
      W_o[7,32] := 0.01371438;
      W_o[7,33] := 0.38752636;
      W_o[7,34] := 0.15796889;
      W_o[7,35] := -0.05519250;
      W_o[7,36] := 0.04871224;
      W_o[7,37] := -0.17531762;
      W_o[7,38] := 0.12556618;
      W_o[7,39] := 0.51951492;
      W_o[8,0] := 0.06394195;
      W_o[8,1] := 0.17076638;
      W_o[8,2] := -0.10039674;
      W_o[8,3] := -0.33651942;
      W_o[8,4] := 0.31007501;
      W_o[8,5] := 0.05197496;
      W_o[8,6] := -0.01656735;
      W_o[8,7] := 0.12790640;
      W_o[8,8] := 0.30033812;
      W_o[8,9] := -0.02012500;
      W_o[8,10] := 0.22443515;
      W_o[8,11] := -0.17770655;
      W_o[8,12] := -0.73770082;
      W_o[8,13] := 0.31852916;
      W_o[8,14] := -0.35518229;
      W_o[8,15] := 0.07199120;
      W_o[8,16] := -0.28111666;
      W_o[8,17] := 0.01000051;
      W_o[8,18] := 0.36765692;
      W_o[8,19] := -0.03547968;
      W_o[8,20] := -0.19686319;
      W_o[8,21] := 0.15272526;
      W_o[8,22] := 0.42476806;
      W_o[8,23] := -0.36033249;
      W_o[8,24] := 1.38535357;
      W_o[8,25] := 1.61054587;
      W_o[8,26] := 0.01937361;
      W_o[8,27] := -0.19785587;
      W_o[8,28] := -0.36753553;
      W_o[8,29] := -0.16174652;
      W_o[8,30] := 0.46827337;
      W_o[8,31] := -0.09923744;
      W_o[8,32] := 0.18555734;
      W_o[8,33] := 0.12179849;
      W_o[8,34] := 1.49276936;
      W_o[8,35] := 0.08704841;
      W_o[8,36] := 0.05555946;
      W_o[8,37] := -0.12351430;
      W_o[8,38] := 0.14559649;
      W_o[8,39] := 0.73714578;
      W_o[9,0] := 0.23104188;
      W_o[9,1] := -0.37553728;
      W_o[9,2] := -0.28727195;
      W_o[9,3] := -0.35031018;
      W_o[9,4] := 0.60829830;
      W_o[9,5] := -0.09552667;
      W_o[9,6] := 0.45592028;
      W_o[9,7] := -0.30415103;
      W_o[9,8] := 0.26670951;
      W_o[9,9] := 0.38333166;
      W_o[9,10] := -0.10408316;
      W_o[9,11] := -0.56295204;
      W_o[9,12] := 0.25366241;
      W_o[9,13] := 0.16823202;
      W_o[9,14] := 0.09202185;
      W_o[9,15] := 0.00952213;
      W_o[9,16] := -0.11405777;
      W_o[9,17] := -0.03855809;
      W_o[9,18] := -0.02253403;
      W_o[9,19] := 0.48154888;
      W_o[9,20] := 0.20891555;
      W_o[9,21] := 0.43464950;
      W_o[9,22] := 0.02325940;
      W_o[9,23] := -0.24670878;
      W_o[9,24] := -0.08609519;
      W_o[9,25] := -0.10266371;
      W_o[9,26] := 0.29583758;
      W_o[9,27] := -0.62991875;
      W_o[9,28] := -0.81162232;
      W_o[9,29] := -1.11133659;
      W_o[9,30] := 0.22002229;
      W_o[9,31] := 0.00901982;
      W_o[9,32] := -0.62355965;
      W_o[9,33] := -0.75333315;
      W_o[9,34] := -1.52598584;
      W_o[9,35] := -0.44686446;
      W_o[9,36] := 0.32879862;
      W_o[9,37] := -0.24673185;
      W_o[9,38] := 0.15742490;
      W_o[9,39] := -0.14049980;
      W_o[10,0] := 0.06652343;
      W_o[10,1] := -0.19470538;
      W_o[10,2] := -0.30487341;
      W_o[10,3] := -0.38069576;
      W_o[10,4] := 0.04057338;
      W_o[10,5] := 0.01880777;
      W_o[10,6] := -0.37193814;
      W_o[10,7] := 0.06555391;
      W_o[10,8] := 0.01233947;
      W_o[10,9] := 0.11164178;
      W_o[10,10] := 0.02777543;
      W_o[10,11] := -0.61474735;
      W_o[10,12] := -0.35695803;
      W_o[10,13] := -0.48645192;
      W_o[10,14] := -0.50885028;
      W_o[10,15] := -0.19305423;
      W_o[10,16] := 0.06526766;
      W_o[10,17] := 0.87165642;
      W_o[10,18] := -0.18345886;
      W_o[10,19] := 0.04411050;
      W_o[10,20] := 0.56275159;
      W_o[10,21] := 0.94484627;
      W_o[10,22] := -0.09950221;
      W_o[10,23] := 0.03454365;
      W_o[10,24] := -0.14066321;
      W_o[10,25] := -0.14744470;
      W_o[10,26] := -0.24545281;
      W_o[10,27] := 0.28469023;
      W_o[10,28] := 0.42433757;
      W_o[10,29] := 0.33172911;
      W_o[10,30] := 0.14359644;
      W_o[10,31] := -0.07731996;
      W_o[10,32] := 0.15873262;
      W_o[10,33] := 0.26325822;
      W_o[10,34] := 0.08210478;
      W_o[10,35] := -0.03535559;
      W_o[10,36] := -0.14255068;
      W_o[10,37] := -0.06271085;
      W_o[10,38] := 0.23752792;
      W_o[10,39] := 0.30014342;
      W_o[11,0] := 0.13154842;
      W_o[11,1] := -0.15394174;
      W_o[11,2] := -0.07008249;
      W_o[11,3] := -0.42792121;
      W_o[11,4] := 0.19656253;
      W_o[11,5] := 0.06030668;
      W_o[11,6] := -0.04454320;
      W_o[11,7] := -0.02605606;
      W_o[11,8] := -0.07528557;
      W_o[11,9] := 0.31813434;
      W_o[11,10] := -0.12571836;
      W_o[11,11] := -0.29872388;
      W_o[11,12] := 0.24146439;
      W_o[11,13] := -0.23881136;
      W_o[11,14] := -0.24915075;
      W_o[11,15] := -0.42647812;
      W_o[11,16] := 0.13256487;
      W_o[11,17] := -0.18015060;
      W_o[11,18] := -0.27864090;
      W_o[11,19] := 0.40441296;
      W_o[11,20] := 0.09091467;
      W_o[11,21] := 0.45153874;
      W_o[11,22] := -0.15325813;
      W_o[11,23] := -0.17464279;
      W_o[11,24] := -0.27042505;
      W_o[11,25] := -0.13127249;
      W_o[11,26] := 0.08290213;
      W_o[11,27] := 0.14768299;
      W_o[11,28] := 0.07636873;
      W_o[11,29] := -0.21547949;
      W_o[11,30] := -0.11796391;
      W_o[11,31] := 0.29416916;
      W_o[11,32] := 0.02105855;
      W_o[11,33] := 0.22922903;
      W_o[11,34] := -1.29468107;
      W_o[11,35] := -0.13968611;
      W_o[11,36] := 0.19066274;
      W_o[11,37] := -0.03171046;
      W_o[11,38] := -0.11227037;
      W_o[11,39] := 0.22209407;
      W_o[12,0] := 1.17421770;
      W_o[12,1] := 0.26429084;
      W_o[12,2] := 0.43585157;
      W_o[12,3] := -0.48518819;
      W_o[12,4] := -0.40976501;
      W_o[12,5] := 0.11100869;
      W_o[12,6] := 0.29647315;
      W_o[12,7] := -0.89749271;
      W_o[12,8] := 1.16584420;
      W_o[12,9] := -0.37191725;
      W_o[12,10] := -0.52895314;
      W_o[12,11] := -0.24108584;
      W_o[12,12] := 0.30931628;
      W_o[12,13] := 0.47943950;
      W_o[12,14] := 0.11668638;
      W_o[12,15] := -0.12159639;
      W_o[12,16] := 0.02150770;
      W_o[12,17] := 0.07519801;
      W_o[12,18] := 0.84063703;
      W_o[12,19] := 0.34892720;
      W_o[12,20] := 0.20678209;
      W_o[12,21] := 0.36131117;
      W_o[12,22] := 0.04332813;
      W_o[12,23] := 0.04741211;
      W_o[12,24] := -0.10370950;
      W_o[12,25] := -0.09042650;
      W_o[12,26] := -0.23766181;
      W_o[12,27] := 0.16998215;
      W_o[12,28] := 0.34490037;
      W_o[12,29] := 0.41028047;
      W_o[12,30] := -0.14397323;
      W_o[12,31] := -0.23349625;
      W_o[12,32] := 0.07464497;
      W_o[12,33] := 0.30076206;
      W_o[12,34] := 0.22199887;
      W_o[12,35] := -0.09407075;
      W_o[12,36] := 0.00139994;
      W_o[12,37] := 0.15236829;
      W_o[12,38] := 0.35288835;
      W_o[12,39] := 0.14806160;
      W_o[13,0] := 0.84261262;
      W_o[13,1] := -0.20696357;
      W_o[13,2] := -0.45374775;
      W_o[13,3] := 0.22621642;
      W_o[13,4] := -0.91789764;
      W_o[13,5] := 0.04173239;
      W_o[13,6] := -0.45060819;
      W_o[13,7] := -0.22334968;
      W_o[13,8] := -0.58925390;
      W_o[13,9] := -0.20284618;
      W_o[13,10] := 0.52314490;
      W_o[13,11] := -0.15634355;
      W_o[13,12] := 0.44538718;
      W_o[13,13] := -0.62631238;
      W_o[13,14] := -0.03795471;
      W_o[13,15] := 0.06832328;
      W_o[13,16] := -0.02699518;
      W_o[13,17] := -0.02816617;
      W_o[13,18] := 0.28338355;
      W_o[13,19] := -0.04717518;
      W_o[13,20] := 0.89906502;
      W_o[13,21] := 0.96378762;
      W_o[13,22] := 0.74177384;
      W_o[13,23] := -0.44595194;
      W_o[13,24] := 1.96999025;
      W_o[13,25] := 1.73697257;
      W_o[13,26] := -0.61652189;
      W_o[13,27] := -0.03462137;
      W_o[13,28] := 0.73489487;
      W_o[13,29] := 0.28480554;
      W_o[13,30] := 0.75282598;
      W_o[13,31] := -0.48566747;
      W_o[13,32] := 0.35734117;
      W_o[13,33] := 0.15278557;
      W_o[13,34] := 1.63127089;
      W_o[13,35] := 0.05970725;
      W_o[13,36] := -0.44636431;
      W_o[13,37] := 0.03125810;
      W_o[13,38] := 0.54704839;
      W_o[13,39] := 0.23915936;
      W_o[14,0] := -0.11508259;
      W_o[14,1] := -0.00742625;
      W_o[14,2] := -0.14038253;
      W_o[14,3] := -0.32177269;
      W_o[14,4] := -0.19025247;
      W_o[14,5] := -0.08554563;
      W_o[14,6] := -0.26530343;
      W_o[14,7] := 0.26199371;
      W_o[14,8] := 0.16477968;
      W_o[14,9] := 0.51352233;
      W_o[14,10] := -0.31731769;
      W_o[14,11] := 0.23585543;
      W_o[14,12] := 0.05539954;
      W_o[14,13] := 0.26555577;
      W_o[14,14] := -0.16365553;
      W_o[14,15] := -0.02076932;
      W_o[14,16] := -0.05403108;
      W_o[14,17] := -0.03535303;
      W_o[14,18] := 0.01533344;
      W_o[14,19] := -0.18407176;
      W_o[14,20] := -1.97634840;
      W_o[14,21] := -0.17147033;
      W_o[14,22] := -0.02276186;
      W_o[14,23] := -0.04953425;
      W_o[14,24] := -0.00544362;
      W_o[14,25] := -0.09639890;
      W_o[14,26] := -0.63560331;
      W_o[14,27] := -0.02849981;
      W_o[14,28] := 0.17682418;
      W_o[14,29] := 0.01651747;
      W_o[14,30] := -0.38656715;
      W_o[14,31] := -0.35627303;
      W_o[14,32] := 0.27490258;
      W_o[14,33] := 0.00227457;
      W_o[14,34] := -0.75013810;
      W_o[14,35] := 0.22019975;
      W_o[14,36] := -0.02764499;
      W_o[14,37] := 0.25156558;
      W_o[14,38] := 0.11675658;
      W_o[14,39] := 0.30231616;
      W_o[15,0] := 0.49589619;
      W_o[15,1] := -0.29518256;
      W_o[15,2] := 0.06588203;
      W_o[15,3] := 0.41961071;
      W_o[15,4] := 0.36646873;
      W_o[15,5] := -0.17609957;
      W_o[15,6] := 0.22730346;
      W_o[15,7] := 0.38059497;
      W_o[15,8] := 0.00410721;
      W_o[15,9] := 0.01834118;
      W_o[15,10] := 0.80458623;
      W_o[15,11] := 0.36880231;
      W_o[15,12] := 0.27834967;
      W_o[15,13] := -0.88198465;
      W_o[15,14] := -1.21522260;
      W_o[15,15] := -0.52633685;
      W_o[15,16] := 0.01724990;
      W_o[15,17] := -0.29456952;
      W_o[15,18] := 0.15491745;
      W_o[15,19] := -0.14392993;
      W_o[15,20] := 0.04712911;
      W_o[15,21] := 1.08945072;
      W_o[15,22] := 0.00751739;
      W_o[15,23] := -0.52356565;
      W_o[15,24] := -0.25086331;
      W_o[15,25] := -0.20301269;
      W_o[15,26] := -0.34148690;
      W_o[15,27] := 0.20905708;
      W_o[15,28] := 0.35473186;
      W_o[15,29] := -0.24059887;
      W_o[15,30] := 0.19723336;
      W_o[15,31] := -0.33502799;
      W_o[15,32] := 0.19524355;
      W_o[15,33] := 0.17764403;
      W_o[15,34] := 0.26448494;
      W_o[15,35] := 0.09686819;
      W_o[15,36] := 0.19879398;
      W_o[15,37] := -0.01141761;
      W_o[15,38] := 0.61595124;
      W_o[15,39] := 1.55151069;
      W_o[16,0] := -0.03918270;
      W_o[16,1] := -0.22132833;
      W_o[16,2] := 0.03094298;
      W_o[16,3] := -0.18334754;
      W_o[16,4] := -0.13022275;
      W_o[16,5] := 0.01883446;
      W_o[16,6] := -0.10264830;
      W_o[16,7] := -0.08231372;
      W_o[16,8] := -0.04199046;
      W_o[16,9] := 0.27921346;
      W_o[16,10] := 0.02591077;
      W_o[16,11] := -0.43003944;
      W_o[16,12] := -0.19622396;
      W_o[16,13] := 0.03951275;
      W_o[16,14] := 0.45676297;
      W_o[16,15] := 0.04330837;
      W_o[16,16] := -0.01354478;
      W_o[16,17] := -0.27774113;
      W_o[16,18] := 0.28355557;
      W_o[16,19] := 0.75274837;
      W_o[16,20] := -0.24724983;
      W_o[16,21] := -0.20417309;
      W_o[16,22] := 0.12291051;
      W_o[16,23] := -0.05004810;
      W_o[16,24] := 0.17314653;
      W_o[16,25] := 0.20202337;
      W_o[16,26] := 0.05929702;
      W_o[16,27] := 0.07103945;
      W_o[16,28] := -0.14921938;
      W_o[16,29] := 0.15395188;
      W_o[16,30] := 0.07721848;
      W_o[16,31] := 0.08066402;
      W_o[16,32] := -0.12877144;
      W_o[16,33] := -0.14650317;
      W_o[16,34] := -0.44100365;
      W_o[16,35] := 0.07829420;
      W_o[16,36] := -0.02766092;
      W_o[16,37] := 0.25472456;
      W_o[16,38] := -0.17556611;
      W_o[16,39] := 0.44761717;
      W_o[17,0] := -0.15512046;
      W_o[17,1] := -0.14749597;
      W_o[17,2] := 0.14577709;
      W_o[17,3] := -0.24457024;
      W_o[17,4] := 0.66728854;
      W_o[17,5] := -0.54898918;
      W_o[17,6] := 0.55137467;
      W_o[17,7] := -0.17406906;
      W_o[17,8] := -0.18214005;
      W_o[17,9] := 0.00611916;
      W_o[17,10] := 0.10385188;
      W_o[17,11] := -0.04477718;
      W_o[17,12] := 0.37598988;
      W_o[17,13] := -0.06295054;
      W_o[17,14] := 0.11274575;
      W_o[17,15] := 0.07089063;
      W_o[17,16] := -0.00096506;
      W_o[17,17] := -0.58720839;
      W_o[17,18] := -0.19919771;
      W_o[17,19] := -0.12993361;
      W_o[17,20] := 0.16244391;
      W_o[17,21] := 1.12817502;
      W_o[17,22] := -0.23536411;
      W_o[17,23] := 0.18415383;
      W_o[17,24] := 0.03566999;
      W_o[17,25] := -0.12391213;
      W_o[17,26] := 0.49041089;
      W_o[17,27] := 0.09547501;
      W_o[17,28] := 0.13685285;
      W_o[17,29] := 0.79314357;
      W_o[17,30] := -0.11405763;
      W_o[17,31] := -0.03408524;
      W_o[17,32] := -0.07211143;
      W_o[17,33] := 0.61566854;
      W_o[17,34] := -0.12214158;
      W_o[17,35] := -0.06288216;
      W_o[17,36] := -0.14356418;
      W_o[17,37] := -0.39446166;
      W_o[17,38] := 0.58293790;
      W_o[17,39] := -0.00185990;
      W_o[18,0] := 0.76430744;
      W_o[18,1] := -0.08611343;
      W_o[18,2] := -0.21489345;
      W_o[18,3] := 0.02633494;
      W_o[18,4] := 0.26816112;
      W_o[18,5] := 0.33768278;
      W_o[18,6] := -0.93157423;
      W_o[18,7] := 0.33818114;
      W_o[18,8] := 0.00433187;
      W_o[18,9] := -0.38866064;
      W_o[18,10] := 0.05605030;
      W_o[18,11] := 0.31501544;
      W_o[18,12] := 0.26311636;
      W_o[18,13] := 0.19155917;
      W_o[18,14] := 0.07760307;
      W_o[18,15] := 0.06348719;
      W_o[18,16] := -0.06047682;
      W_o[18,17] := 0.04179845;
      W_o[18,18] := -0.07208342;
      W_o[18,19] := -0.55079585;
      W_o[18,20] := -0.58557802;
      W_o[18,21] := -0.12302866;
      W_o[18,22] := -0.06828116;
      W_o[18,23] := -0.27328676;
      W_o[18,24] := -0.02747243;
      W_o[18,25] := -0.23128007;
      W_o[18,26] := 0.45590901;
      W_o[18,27] := 0.62222111;
      W_o[18,28] := -0.22750355;
      W_o[18,29] := -0.68637496;
      W_o[18,30] := 0.02868916;
      W_o[18,31] := -0.81999731;
      W_o[18,32] := 0.14697376;
      W_o[18,33] := -0.01794586;
      W_o[18,34] := -0.70916694;
      W_o[18,35] := 0.42292288;
      W_o[18,36] := -0.45709130;
      W_o[18,37] := 0.86393505;
      W_o[18,38] := -0.07340389;
      W_o[18,39] := -0.15890661;
      W_o[19,0] := 0.29933581;
      W_o[19,1] := -0.24707638;
      W_o[19,2] := 0.01626565;
      W_o[19,3] := 0.12035257;
      W_o[19,4] := -0.37100369;
      W_o[19,5] := -0.16028123;
      W_o[19,6] := 0.52533126;
      W_o[19,7] := -0.45668989;
      W_o[19,8] := 0.01525003;
      W_o[19,9] := -1.26570213;
      W_o[19,10] := 1.04233599;
      W_o[19,11] := 0.21994767;
      W_o[19,12] := 0.43801033;
      W_o[19,13] := -0.07208458;
      W_o[19,14] := -0.10423371;
      W_o[19,15] := 0.00277623;
      W_o[19,16] := 0.17693250;
      W_o[19,17] := -0.49376789;
      W_o[19,18] := -0.31587574;
      W_o[19,19] := -1.32079959;
      W_o[19,20] := -0.11124548;
      W_o[19,21] := 0.18118487;
      W_o[19,22] := 0.20466328;
      W_o[19,23] := 0.27020007;
      W_o[19,24] := 1.90587401;
      W_o[19,25] := 2.08124018;
      W_o[19,26] := 0.13651226;
      W_o[19,27] := 0.32710886;
      W_o[19,28] := 0.41084310;
      W_o[19,29] := 0.66397214;
      W_o[19,30] := 0.30322510;
      W_o[19,31] := 0.17320575;
      W_o[19,32] := -0.12189152;
      W_o[19,33] := 0.31796196;
      W_o[19,34] := -0.16206127;
      W_o[19,35] := -0.32837775;
      W_o[19,36] := 0.09268205;
      W_o[19,37] := -0.41775760;
      W_o[19,38] := -0.08859571;
      W_o[19,39] := -0.03335560;
      W_o[20,0] := 0.13922459;
      W_o[20,1] := -2.20053363;
      W_o[20,2] := 0.00205416;
      W_o[20,3] := 0.21276508;
      W_o[20,4] := 0.27908573;
      W_o[20,5] := 0.01135337;
      W_o[20,6] := 0.01100084;
      W_o[20,7] := 0.44203964;
      W_o[20,8] := -0.68097985;
      W_o[20,9] := -0.37706792;
      W_o[20,10] := 0.35476449;
      W_o[20,11] := -0.60206777;
      W_o[20,12] := 0.08790465;
      W_o[20,13] := -0.36102074;
      W_o[20,14] := -0.01076331;
      W_o[20,15] := 0.16372751;
      W_o[20,16] := -0.14292030;
      W_o[20,17] := -0.03609731;
      W_o[20,18] := -0.24819231;
      W_o[20,19] := 0.02868344;
      W_o[20,20] := 0.09508435;
      W_o[20,21] := 0.10375975;
      W_o[20,22] := -0.13606212;
      W_o[20,23] := -0.75565112;
      W_o[20,24] := 1.13532817;
      W_o[20,25] := 0.80740219;
      W_o[20,26] := 0.26416770;
      W_o[20,27] := 0.49109095;
      W_o[20,28] := -0.13837487;
      W_o[20,29] := -0.17751533;
      W_o[20,30] := -0.20410518;
      W_o[20,31] := -0.19428243;
      W_o[20,32] := 0.01627112;
      W_o[20,33] := 0.09347031;
      W_o[20,34] := 0.24445274;
      W_o[20,35] := -0.21534006;
      W_o[20,36] := 0.06837694;
      W_o[20,37] := -0.24603793;
      W_o[20,38] := 0.09559119;
      W_o[20,39] := 0.09811132;
      W_o[21,0] := -0.10988021;
      W_o[21,1] := 0.24835177;
      W_o[21,2] := -0.44709471;
      W_o[21,3] := -0.23855081;
      W_o[21,4] := -0.05993883;
      W_o[21,5] := 0.05487840;
      W_o[21,6] := 0.30802393;
      W_o[21,7] := 0.20565377;
      W_o[21,8] := 0.01227701;
      W_o[21,9] := 0.17216517;
      W_o[21,10] := -0.24846844;
      W_o[21,11] := -0.05311755;
      W_o[21,12] := 0.14346336;
      W_o[21,13] := -0.01710485;
      W_o[21,14] := 0.01053591;
      W_o[21,15] := -0.30249557;
      W_o[21,16] := -0.03592461;
      W_o[21,17] := -0.01890021;
      W_o[21,18] := -0.18794870;
      W_o[21,19] := -0.04519326;
      W_o[21,20] := -0.22630790;
      W_o[21,21] := 0.82546812;
      W_o[21,22] := 0.16347410;
      W_o[21,23] := 0.34241235;
      W_o[21,24] := 0.78471315;
      W_o[21,25] := 0.11163335;
      W_o[21,26] := -0.04875318;
      W_o[21,27] := -0.10537915;
      W_o[21,28] := 0.35267621;
      W_o[21,29] := 0.14096136;
      W_o[21,30] := 0.19667439;
      W_o[21,31] := -0.05898595;
      W_o[21,32] := -0.17870322;
      W_o[21,33] := 0.03267650;
      W_o[21,34] := -0.40305266;
      W_o[21,35] := -0.04123265;
      W_o[21,36] := 0.96496969;
      W_o[21,37] := 0.20428683;
      W_o[21,38] := 0.35514468;
      W_o[21,39] := 0.03118325;
      W_o[22,0] := 0.41157860;
      W_o[22,1] := -0.32734281;
      W_o[22,2] := 0.15231930;
      W_o[22,3] := -0.15504754;
      W_o[22,4] := 0.16780476;
      W_o[22,5] := 0.61459172;
      W_o[22,6] := 0.05332777;
      W_o[22,7] := -0.03754049;
      W_o[22,8] := -0.17407671;
      W_o[22,9] := -0.16621305;
      W_o[22,10] := 0.10367353;
      W_o[22,11] := -0.12657513;
      W_o[22,12] := -0.26324561;
      W_o[22,13] := -0.22081058;
      W_o[22,14] := -0.46252978;
      W_o[22,15] := -0.48273844;
      W_o[22,16] := -0.56322485;
      W_o[22,17] := -0.06665193;
      W_o[22,18] := 1.14411294;
      W_o[22,19] := -0.33045414;
      W_o[22,20] := -0.05424431;
      W_o[22,21] := 0.34366548;
      W_o[22,22] := 0.13654912;
      W_o[22,23] := 0.48519036;
      W_o[22,24] := 0.16035570;
      W_o[22,25] := 0.11601855;
      W_o[22,26] := -0.51481938;
      W_o[22,27] := 0.09939534;
      W_o[22,28] := -0.30302757;
      W_o[22,29] := 0.27184495;
      W_o[22,30] := 0.14510697;
      W_o[22,31] := 0.07548800;
      W_o[22,32] := 0.11845539;
      W_o[22,33] := 0.00411626;
      W_o[22,34] := 0.21212496;
      W_o[22,35] := 0.03143089;
      W_o[22,36] := 0.21655953;
      W_o[22,37] := 0.34552658;
      W_o[22,38] := 0.08682747;
      W_o[22,39] := 0.58460540;
      W_o[23,0] := 0.11161003;
      W_o[23,1] := 0.24242438;
      W_o[23,2] := -0.06118851;
      W_o[23,3] := 0.02698644;
      W_o[23,4] := 0.25399089;
      W_o[23,5] := 0.52320135;
      W_o[23,6] := -0.80968732;
      W_o[23,7] := 0.31103149;
      W_o[23,8] := -0.01249438;
      W_o[23,9] := 0.58440495;
      W_o[23,10] := -0.85927993;
      W_o[23,11] := -0.35480243;
      W_o[23,12] := -0.12797940;
      W_o[23,13] := 0.12250131;
      W_o[23,14] := -0.03641031;
      W_o[23,15] := 0.09557875;
      W_o[23,16] := 0.06768897;
      W_o[23,17] := 0.07494175;
      W_o[23,18] := 0.12114435;
      W_o[23,19] := 0.04627066;
      W_o[23,20] := -0.22720096;
      W_o[23,21] := 0.18305890;
      W_o[23,22] := -0.22875017;
      W_o[23,23] := 0.47580439;
      W_o[23,24] := -0.21235433;
      W_o[23,25] := -0.20607333;
      W_o[23,26] := -0.24356085;
      W_o[23,27] := 0.49107108;
      W_o[23,28] := -0.05528429;
      W_o[23,29] := -0.22709295;
      W_o[23,30] := -0.21775801;
      W_o[23,31] := 0.04588168;
      W_o[23,32] := -0.02398799;
      W_o[23,33] := -0.03821435;
      W_o[23,34] := -0.01893564;
      W_o[23,35] := -0.01355231;
      W_o[23,36] := -0.09647775;
      W_o[23,37] := -0.08327264;
      W_o[23,38] := -0.10612083;
      W_o[23,39] := 0.02147446;
      W_o[24,0] := 0.92537642;
      W_o[24,1] := -0.01338725;
      W_o[24,2] := -0.29871222;
      W_o[24,3] := 0.36259899;
      W_o[24,4] := 0.29513517;
      W_o[24,5] := -0.12575051;
      W_o[24,6] := -0.00142940;
      W_o[24,7] := -0.12991576;
      W_o[24,8] := -0.39490813;
      W_o[24,9] := 0.25243637;
      W_o[24,10] := -0.01860771;
      W_o[24,11] := -0.39029965;
      W_o[24,12] := 0.34209472;
      W_o[24,13] := -0.69206321;
      W_o[24,14] := 0.01371827;
      W_o[24,15] := -0.03120338;
      W_o[24,16] := 0.08943855;
      W_o[24,17] := 0.00575395;
      W_o[24,18] := -0.05534322;
      W_o[24,19] := -0.13040026;
      W_o[24,20] := 0.12296753;
      W_o[24,21] := -0.49935907;
      W_o[24,22] := -0.33874360;
      W_o[24,23] := -0.54052353;
      W_o[24,24] := 1.64606535;
      W_o[24,25] := 1.50577116;
      W_o[24,26] := -0.29378295;
      W_o[24,27] := 0.70552373;
      W_o[24,28] := -0.84343106;
      W_o[24,29] := 0.64516312;
      W_o[24,30] := -0.53515697;
      W_o[24,31] := -0.02786028;
      W_o[24,32] := 0.06958819;
      W_o[24,33] := 0.09729471;
      W_o[24,34] := 0.74627382;
      W_o[24,35] := 0.67337501;
      W_o[24,36] := -0.10799170;
      W_o[24,37] := 0.99782586;
      W_o[24,38] := -0.04200582;
      W_o[24,39] := 0.22245386;
      W_o[25,0] := -0.07363706;
      W_o[25,1] := -0.28953281;
      W_o[25,2] := -0.02809429;
      W_o[25,3] := 0.08961703;
      W_o[25,4] := 0.07100378;
      W_o[25,5] := 0.00981856;
      W_o[25,6] := 0.05789235;
      W_o[25,7] := -0.11700267;
      W_o[25,8] := 0.13359351;
      W_o[25,9] := -0.30955857;
      W_o[25,10] := 0.04413471;
      W_o[25,11] := 0.19343543;
      W_o[25,12] := 0.72226489;
      W_o[25,13] := 0.11818234;
      W_o[25,14] := -0.30286118;
      W_o[25,15] := -0.90309602;
      W_o[25,16] := 0.01062219;
      W_o[25,17] := -0.32118207;
      W_o[25,18] := -0.07703356;
      W_o[25,19] := -0.12701164;
      W_o[25,20] := -0.14186306;
      W_o[25,21] := 0.26098636;
      W_o[25,22] := 0.06865875;
      W_o[25,23] := -0.19780582;
      W_o[25,24] := 0.26296347;
      W_o[25,25] := 0.19853988;
      W_o[25,26] := 0.03239297;
      W_o[25,27] := -0.29850340;
      W_o[25,28] := -0.26168373;
      W_o[25,29] := -0.09161076;
      W_o[25,30] := 0.04232042;
      W_o[25,31] := -0.16418776;
      W_o[25,32] := 0.24403407;
      W_o[25,33] := 0.08130822;
      W_o[25,34] := -1.18890846;
      W_o[25,35] := 0.01663818;
      W_o[25,36] := -0.04253452;
      W_o[25,37] := 0.33604178;
      W_o[25,38] := 0.01961804;
      W_o[25,39] := 0.04668290;
      W_o[26,0] := -0.05728961;
      W_o[26,1] := -0.04979565;
      W_o[26,2] := -0.02092489;
      W_o[26,3] := -0.03078631;
      W_o[26,4] := -0.16870457;
      W_o[26,5] := -0.10186446;
      W_o[26,6] := -0.10564874;
      W_o[26,7] := -0.06154874;
      W_o[26,8] := 0.00327657;
      W_o[26,9] := -0.00514480;
      W_o[26,10] := 0.01865643;
      W_o[26,11] := 0.06774835;
      W_o[26,12] := 0.00966269;
      W_o[26,13] := -0.02320647;
      W_o[26,14] := -0.00139932;
      W_o[26,15] := -0.12217309;
      W_o[26,16] := -0.02373873;
      W_o[26,17] := 0.01413365;
      W_o[26,18] := 1.74683726;
      W_o[26,19] := 0.00071617;
      W_o[26,20] := -0.09387178;
      W_o[26,21] := -0.16163847;
      W_o[26,22] := -0.07811227;
      W_o[26,23] := 0.12433856;
      W_o[26,24] := 0.40757918;
      W_o[26,25] := 0.23269270;
      W_o[26,26] := 0.06876845;
      W_o[26,27] := 0.19421263;
      W_o[26,28] := 0.01647574;
      W_o[26,29] := 0.03276436;
      W_o[26,30] := -0.11340243;
      W_o[26,31] := -0.01652885;
      W_o[26,32] := -0.04143284;
      W_o[26,33] := -0.00182136;
      W_o[26,34] := -0.31087825;
      W_o[26,35] := -0.28638926;
      W_o[26,36] := -0.01335451;
      W_o[26,37] := -0.27111626;
      W_o[26,38] := -0.00584449;
      W_o[26,39] := 1.61455750;
      W_o[27,0] := 0.14007252;
      W_o[27,1] := -0.11251914;
      W_o[27,2] := -0.01313373;
      W_o[27,3] := -0.08391760;
      W_o[27,4] := -0.07205343;
      W_o[27,5] := -0.21357708;
      W_o[27,6] := 0.08899514;
      W_o[27,7] := -0.12406176;
      W_o[27,8] := 0.16971087;
      W_o[27,9] := 0.42553920;
      W_o[27,10] := 0.09811529;
      W_o[27,11] := -1.13219488;
      W_o[27,12] := 0.25516251;
      W_o[27,13] := 0.08068778;
      W_o[27,14] := 0.16564816;
      W_o[27,15] := -0.44411266;
      W_o[27,16] := -0.05831531;
      W_o[27,17] := -0.41473165;
      W_o[27,18] := -0.03482730;
      W_o[27,19] := -0.05169702;
      W_o[27,20] := -0.11636675;
      W_o[27,21] := 0.04912658;
      W_o[27,22] := -0.11369362;
      W_o[27,23] := -0.08044525;
      W_o[27,24] := 1.32685113;
      W_o[27,25] := 1.29689372;
      W_o[27,26] := 0.17168416;
      W_o[27,27] := 0.01350123;
      W_o[27,28] := 0.04110165;
      W_o[27,29] := -0.66268092;
      W_o[27,30] := -0.13212320;
      W_o[27,31] := -0.01355234;
      W_o[27,32] := -0.26603335;
      W_o[27,33] := -0.43971109;
      W_o[27,34] := 0.47377747;
      W_o[27,35] := -0.08899359;
      W_o[27,36] := 0.05804361;
      W_o[27,37] := -0.01794386;
      W_o[27,38] := -0.16820285;
      W_o[27,39] := 0.37586251;
      W_o[28,0] := -0.31159109;
      W_o[28,1] := -0.09061144;
      W_o[28,2] := -0.01196734;
      W_o[28,3] := -0.62155133;
      W_o[28,4] := 0.36044863;
      W_o[28,5] := -0.00623550;
      W_o[28,6] := 0.33896664;
      W_o[28,7] := 0.45510116;
      W_o[28,8] := -0.66868389;
      W_o[28,9] := 0.28924412;
      W_o[28,10] := 0.39494881;
      W_o[28,11] := 0.06208984;
      W_o[28,12] := -0.07699963;
      W_o[28,13] := 0.47504538;
      W_o[28,14] := -0.05790047;
      W_o[28,15] := -0.08396290;
      W_o[28,16] := -0.49277100;
      W_o[28,17] := 0.26957941;
      W_o[28,18] := 0.11747041;
      W_o[28,19] := 0.48421782;
      W_o[28,20] := -0.05510560;
      W_o[28,21] := -0.27798435;
      W_o[28,22] := -0.08301591;
      W_o[28,23] := -0.08954213;
      W_o[28,24] := 1.51879895;
      W_o[28,25] := 2.18036342;
      W_o[28,26] := 0.14471918;
      W_o[28,27] := 0.66814166;
      W_o[28,28] := -0.34997442;
      W_o[28,29] := -0.11917944;
      W_o[28,30] := -0.16639628;
      W_o[28,31] := 0.10294037;
      W_o[28,32] := -0.36679235;
      W_o[28,33] := -0.27575570;
      W_o[28,34] := 0.14579554;
      W_o[28,35] := -0.24746421;
      W_o[28,36] := -0.13615337;
      W_o[28,37] := -0.41702220;
      W_o[28,38] := 0.00291938;
      W_o[28,39] := -0.06635363;
      W_o[29,0] := 0.25321370;
      W_o[29,1] := -0.28984985;
      W_o[29,2] := 0.14680482;
      W_o[29,3] := -0.22666040;
      W_o[29,4] := 0.17676389;
      W_o[29,5] := 0.64302081;
      W_o[29,6] := -0.20920402;
      W_o[29,7] := 0.13273127;
      W_o[29,8] := 0.13646045;
      W_o[29,9] := -0.51564175;
      W_o[29,10] := -0.46837211;
      W_o[29,11] := -0.10658596;
      W_o[29,12] := 0.34777194;
      W_o[29,13] := 0.00625758;
      W_o[29,14] := 0.02718482;
      W_o[29,15] := -0.03930616;
      W_o[29,16] := 0.14963950;
      W_o[29,17] := 0.02233061;
      W_o[29,18] := 0.96453893;
      W_o[29,19] := 0.14056733;
      W_o[29,20] := -0.46394807;
      W_o[29,21] := 0.52843809;
      W_o[29,22] := -0.14849740;
      W_o[29,23] := 1.63552296;
      W_o[29,24] := 0.13075085;
      W_o[29,25] := 0.15701653;
      W_o[29,26] := -0.09133709;
      W_o[29,27] := 0.43826416;
      W_o[29,28] := -0.04762744;
      W_o[29,29] := 0.02618933;
      W_o[29,30] := -0.15002266;
      W_o[29,31] := 0.15962145;
      W_o[29,32] := 0.04751491;
      W_o[29,33] := -0.34306863;
      W_o[29,34] := -0.35635781;
      W_o[29,35] := 0.05356752;
      W_o[29,36] := 0.06037952;
      W_o[29,37] := 0.03712659;
      W_o[29,38] := 0.02771435;
      W_o[29,39] := 0.69680142;
      W_o[30,0] := -0.27389616;
      W_o[30,1] := -0.33204398;
      W_o[30,2] := 0.21435702;
      W_o[30,3] := -0.19798888;
      W_o[30,4] := -0.09623803;
      W_o[30,5] := 0.87759387;
      W_o[30,6] := 0.46116766;
      W_o[30,7] := -0.01188846;
      W_o[30,8] := -0.17874885;
      W_o[30,9] := 0.09584995;
      W_o[30,10] := 0.38583899;
      W_o[30,11] := -0.70979095;
      W_o[30,12] := 0.12901115;
      W_o[30,13] := -0.28334385;
      W_o[30,14] := -0.35588500;
      W_o[30,15] := -1.42531514;
      W_o[30,16] := -0.59441978;
      W_o[30,17] := 0.14774412;
      W_o[30,18] := 0.18592946;
      W_o[30,19] := 0.93774903;
      W_o[30,20] := 0.17501442;
      W_o[30,21] := 0.40653196;
      W_o[30,22] := -0.03565990;
      W_o[30,23] := 0.01427438;
      W_o[30,24] := 0.00282043;
      W_o[30,25] := 0.10861620;
      W_o[30,26] := 0.04156169;
      W_o[30,27] := -0.05955997;
      W_o[30,28] := 0.23415500;
      W_o[30,29] := -0.10069150;
      W_o[30,30] := 0.12966040;
      W_o[30,31] := 0.20069182;
      W_o[30,32] := 0.13809177;
      W_o[30,33] := 0.33505166;
      W_o[30,34] := 0.40418807;
      W_o[30,35] := -0.14144862;
      W_o[30,36] := 0.07608719;
      W_o[30,37] := -0.11019205;
      W_o[30,38] := 0.47189629;
      W_o[30,39] := 0.06401872;
      W_o[31,0] := -0.15408427;
      W_o[31,1] := -0.35604635;
      W_o[31,2] := 0.14469552;
      W_o[31,3] := 0.01747640;
      W_o[31,4] := -0.10457193;
      W_o[31,5] := -0.03063329;
      W_o[31,6] := 0.22982945;
      W_o[31,7] := -0.18897052;
      W_o[31,8] := -0.10540372;
      W_o[31,9] := -0.02604771;
      W_o[31,10] := -0.00690281;
      W_o[31,11] := -0.60990834;
      W_o[31,12] := 0.31482366;
      W_o[31,13] := 0.03766366;
      W_o[31,14] := -0.04685820;
      W_o[31,15] := 0.21878938;
      W_o[31,16] := -0.13059433;
      W_o[31,17] := 0.06215651;
      W_o[31,18] := -0.08466318;
      W_o[31,19] := -0.53358144;
      W_o[31,20] := -0.04495485;
      W_o[31,21] := -0.19969423;
      W_o[31,22] := 0.11028804;
      W_o[31,23] := 0.14346430;
      W_o[31,24] := 0.34848404;
      W_o[31,25] := 0.01787481;
      W_o[31,26] := -0.01638452;
      W_o[31,27] := -0.05403485;
      W_o[31,28] := -0.02076081;
      W_o[31,29] := 0.63390154;
      W_o[31,30] := 0.08677601;
      W_o[31,31] := 0.00503407;
      W_o[31,32] := 0.11718934;
      W_o[31,33] := -0.02121959;
      W_o[31,34] := -0.82473320;
      W_o[31,35] := 0.33167773;
      W_o[31,36] := -0.00783546;
      W_o[31,37] := 0.39109421;
      W_o[31,38] := 0.27141920;
      W_o[31,39] := 0.05769989;
      R_i[0,0] := -0.45433718;
      R_i[0,1] := 0.04381683;
      R_i[0,2] := 0.06890769;
      R_i[0,3] := 0.29077119;
      R_i[0,4] := 0.36511230;
      R_i[0,5] := 0.71392870;
      R_i[0,6] := -0.57234347;
      R_i[0,7] := 0.08876300;
      R_i[0,8] := 1.04849303;
      R_i[0,9] := 0.47379592;
      R_i[0,10] := 0.81098163;
      R_i[0,11] := -1.16598749;
      R_i[0,12] := -0.15472579;
      R_i[0,13] := -0.10207538;
      R_i[0,14] := -0.02121414;
      R_i[0,15] := -0.51939249;
      R_i[0,16] := -0.28122181;
      R_i[0,17] := 1.61604273;
      R_i[0,18] := -0.04420009;
      R_i[0,19] := 0.70076549;
      R_i[0,20] := 0.33963588;
      R_i[0,21] := 0.52128637;
      R_i[0,22] := 0.16769774;
      R_i[0,23] := -0.01815144;
      R_i[0,24] := 0.26494589;
      R_i[0,25] := -0.31607488;
      R_i[0,26] := 0.43812805;
      R_i[0,27] := -0.78570491;
      R_i[0,28] := 0.20476782;
      R_i[0,29] := -0.48682672;
      R_i[0,30] := 0.40167305;
      R_i[0,31] := 0.31006321;
      R_i[1,0] := -0.13692026;
      R_i[1,1] := -0.24063189;
      R_i[1,2] := 0.22683647;
      R_i[1,3] := -0.18372364;
      R_i[1,4] := -0.23403043;
      R_i[1,5] := -0.09768691;
      R_i[1,6] := 0.39038301;
      R_i[1,7] := 0.11476605;
      R_i[1,8] := 0.08316614;
      R_i[1,9] := 0.35416487;
      R_i[1,10] := -0.18735920;
      R_i[1,11] := -0.31722569;
      R_i[1,12] := 0.20257886;
      R_i[1,13] := 0.10904857;
      R_i[1,14] := -0.11465105;
      R_i[1,15] := 0.33582023;
      R_i[1,16] := 0.06933430;
      R_i[1,17] := 0.21575241;
      R_i[1,18] := 0.41760844;
      R_i[1,19] := -0.03354438;
      R_i[1,20] := 0.11415303;
      R_i[1,21] := -0.70651364;
      R_i[1,22] := -0.08349572;
      R_i[1,23] := 0.28775278;
      R_i[1,24] := -1.60818112;
      R_i[1,25] := -0.10913862;
      R_i[1,26] := 0.23515795;
      R_i[1,27] := -0.07737515;
      R_i[1,28] := 0.05925220;
      R_i[1,29] := 0.36150515;
      R_i[1,30] := -0.12552686;
      R_i[1,31] := 0.50926840;
      R_i[2,0] := -0.05818795;
      R_i[2,1] := -0.28729683;
      R_i[2,2] := 0.45500574;
      R_i[2,3] := 0.12803800;
      R_i[2,4] := -0.02028978;
      R_i[2,5] := -0.06158508;
      R_i[2,6] := 0.06124555;
      R_i[2,7] := 0.07490601;
      R_i[2,8] := 0.28868538;
      R_i[2,9] := 0.30742335;
      R_i[2,10] := 0.31020564;
      R_i[2,11] := -0.40941274;
      R_i[2,12] := -0.52057606;
      R_i[2,13] := 0.34527487;
      R_i[2,14] := -0.25903773;
      R_i[2,15] := 0.57880473;
      R_i[2,16] := 0.04028931;
      R_i[2,17] := 0.77455544;
      R_i[2,18] := 0.05028503;
      R_i[2,19] := -0.31733224;
      R_i[2,20] := 0.60684431;
      R_i[2,21] := -0.56939471;
      R_i[2,22] := 0.21272865;
      R_i[2,23] := -0.22903784;
      R_i[2,24] := -1.24987829;
      R_i[2,25] := 0.00797278;
      R_i[2,26] := 0.17857899;
      R_i[2,27] := -0.06947280;
      R_i[2,28] := -0.26714545;
      R_i[2,29] := -0.10779256;
      R_i[2,30] := 0.06115891;
      R_i[2,31] := 0.26452520;
      R_i[3,0] := 0.39931396;
      R_i[3,1] := 1.15073752;
      R_i[3,2] := -0.10358425;
      R_i[3,3] := 0.67767721;
      R_i[3,4] := 0.31121764;
      R_i[3,5] := -0.28151646;
      R_i[3,6] := 0.05488693;
      R_i[3,7] := -0.02619875;
      R_i[3,8] := -0.26502672;
      R_i[3,9] := 0.26960725;
      R_i[3,10] := -0.09923731;
      R_i[3,11] := 0.50374937;
      R_i[3,12] := -0.23172866;
      R_i[3,13] := -0.63132286;
      R_i[3,14] := -0.35142949;
      R_i[3,15] := -0.36325392;
      R_i[3,16] := 0.49311674;
      R_i[3,17] := -0.10561612;
      R_i[3,18] := -0.87026656;
      R_i[3,19] := 0.38533220;
      R_i[3,20] := 0.49307376;
      R_i[3,21] := -0.01616472;
      R_i[3,22] := 0.58301890;
      R_i[3,23] := -0.91731554;
      R_i[3,24] := 0.74190807;
      R_i[3,25] := -0.81879312;
      R_i[3,26] := 0.07494108;
      R_i[3,27] := 0.11778155;
      R_i[3,28] := -0.41089514;
      R_i[3,29] := 0.07875212;
      R_i[3,30] := 0.63496423;
      R_i[3,31] := -0.49545658;
      R_i[4,0] := 0.18378885;
      R_i[4,1] := -0.28184643;
      R_i[4,2] := -0.32651404;
      R_i[4,3] := -1.46459544;
      R_i[4,4] := -0.85016924;
      R_i[4,5] := -0.23196834;
      R_i[4,6] := 1.07934105;
      R_i[4,7] := -0.33986455;
      R_i[4,8] := -1.04742646;
      R_i[4,9] := 0.12250885;
      R_i[4,10] := 0.30320376;
      R_i[4,11] := 0.03586194;
      R_i[4,12] := 0.16321847;
      R_i[4,13] := -0.84031409;
      R_i[4,14] := -0.30363435;
      R_i[4,15] := -0.89096338;
      R_i[4,16] := -0.41343698;
      R_i[4,17] := 0.74893546;
      R_i[4,18] := 0.20611791;
      R_i[4,19] := 0.21939717;
      R_i[4,20] := 0.74230492;
      R_i[4,21] := -0.07196729;
      R_i[4,22] := -0.09799778;
      R_i[4,23] := -0.51248717;
      R_i[4,24] := 1.20486891;
      R_i[4,25] := 0.02356974;
      R_i[4,26] := 0.12652595;
      R_i[4,27] := 1.98098385;
      R_i[4,28] := -0.52964228;
      R_i[4,29] := 0.35606074;
      R_i[4,30] := 0.26468128;
      R_i[4,31] := 0.50841063;
      R_i[5,0] := -0.16141868;
      R_i[5,1] := 0.42481518;
      R_i[5,2] := -0.11765660;
      R_i[5,3] := 0.37742898;
      R_i[5,4] := -0.10233248;
      R_i[5,5] := -0.27804697;
      R_i[5,6] := 0.30110398;
      R_i[5,7] := 0.10596237;
      R_i[5,8] := 0.16512184;
      R_i[5,9] := -0.00419395;
      R_i[5,10] := -0.27078024;
      R_i[5,11] := 0.02054108;
      R_i[5,12] := -0.16205336;
      R_i[5,13] := -0.18527851;
      R_i[5,14] := 0.43905500;
      R_i[5,15] := -0.17345172;
      R_i[5,16] := 0.00580292;
      R_i[5,17] := -0.24766308;
      R_i[5,18] := -0.08646183;
      R_i[5,19] := 0.36573070;
      R_i[5,20] := 0.25471163;
      R_i[5,21] := -0.37055936;
      R_i[5,22] := 0.69699669;
      R_i[5,23] := -0.32280406;
      R_i[5,24] := 0.51599389;
      R_i[5,25] := 0.09720933;
      R_i[5,26] := 0.73423731;
      R_i[5,27] := -0.14514761;
      R_i[5,28] := 0.07095706;
      R_i[5,29] := 0.26992759;
      R_i[5,30] := 0.24137810;
      R_i[5,31] := 0.20172344;
      R_i[6,0] := 0.30367762;
      R_i[6,1] := -0.47776160;
      R_i[6,2] := -0.37913454;
      R_i[6,3] := 0.39747033;
      R_i[6,4] := -0.56866300;
      R_i[6,5] := -0.12954362;
      R_i[6,6] := -0.97472411;
      R_i[6,7] := 0.28027597;
      R_i[6,8] := 0.57420611;
      R_i[6,9] := -0.37255341;
      R_i[6,10] := -0.44898850;
      R_i[6,11] := 0.37070736;
      R_i[6,12] := 0.32810879;
      R_i[6,13] := 0.49652654;
      R_i[6,14] := 0.10154562;
      R_i[6,15] := -0.42494139;
      R_i[6,16] := 0.53713739;
      R_i[6,17] := -0.15384643;
      R_i[6,18] := 0.06196346;
      R_i[6,19] := -1.25819671;
      R_i[6,20] := 0.08705294;
      R_i[6,21] := 0.21311060;
      R_i[6,22] := 0.06580897;
      R_i[6,23] := 0.21626072;
      R_i[6,24] := -0.09428816;
      R_i[6,25] := 0.24361600;
      R_i[6,26] := 0.20728236;
      R_i[6,27] := -0.00100759;
      R_i[6,28] := 0.43091920;
      R_i[6,29] := -0.28887641;
      R_i[6,30] := -0.02350107;
      R_i[6,31] := -0.26930115;
      R_i[7,0] := -0.36902297;
      R_i[7,1] := 0.53722495;
      R_i[7,2] := 0.22628103;
      R_i[7,3] := -0.50461161;
      R_i[7,4] := 0.13517481;
      R_i[7,5] := 0.24313395;
      R_i[7,6] := -0.06336830;
      R_i[7,7] := -0.87224251;
      R_i[7,8] := 0.31494582;
      R_i[7,9] := 0.56106687;
      R_i[7,10] := -0.50384265;
      R_i[7,11] := -0.57320881;
      R_i[7,12] := -0.76926386;
      R_i[7,13] := -0.09765702;
      R_i[7,14] := -0.06975676;
      R_i[7,15] := 0.31892934;
      R_i[7,16] := -0.06996145;
      R_i[7,17] := 0.07684433;
      R_i[7,18] := 0.52881980;
      R_i[7,19] := -0.12767319;
      R_i[7,20] := 0.40447325;
      R_i[7,21] := -0.03331390;
      R_i[7,22] := -0.31306756;
      R_i[7,23] := -0.81669295;
      R_i[7,24] := -0.40777335;
      R_i[7,25] := -0.26863009;
      R_i[7,26] := -0.15568426;
      R_i[7,27] := -0.35343477;
      R_i[7,28] := -0.81822574;
      R_i[7,29] := 0.58622450;
      R_i[7,30] := 0.43811530;
      R_i[7,31] := -0.13610241;
      R_i[8,0] := 0.13995494;
      R_i[8,1] := 0.18966211;
      R_i[8,2] := -0.13668501;
      R_i[8,3] := -0.48719549;
      R_i[8,4] := 0.00925596;
      R_i[8,5] := -0.41893780;
      R_i[8,6] := 0.17539361;
      R_i[8,7] := 0.03431849;
      R_i[8,8] := 0.48571968;
      R_i[8,9] := 0.13743351;
      R_i[8,10] := -0.49978310;
      R_i[8,11] := -0.51658124;
      R_i[8,12] := -0.18935153;
      R_i[8,13] := -0.06984410;
      R_i[8,14] := -0.40678748;
      R_i[8,15] := 0.29402977;
      R_i[8,16] := -0.22782041;
      R_i[8,17] := -0.07687777;
      R_i[8,18] := -0.13222699;
      R_i[8,19] := -1.02457535;
      R_i[8,20] := 0.10192242;
      R_i[8,21] := -0.15518960;
      R_i[8,22] := 0.64550126;
      R_i[8,23] := 0.15165904;
      R_i[8,24] := 0.04112607;
      R_i[8,25] := -0.41499722;
      R_i[8,26] := 0.15730077;
      R_i[8,27] := -0.06758537;
      R_i[8,28] := -0.21931611;
      R_i[8,29] := 0.35440147;
      R_i[8,30] := 0.42760614;
      R_i[8,31] := -0.37057987;
      R_i[9,0] := -0.56370252;
      R_i[9,1] := 0.68367869;
      R_i[9,2] := -0.74821293;
      R_i[9,3] := -0.29154259;
      R_i[9,4] := 0.24524473;
      R_i[9,5] := 0.31957385;
      R_i[9,6] := 0.21675618;
      R_i[9,7] := -0.44607636;
      R_i[9,8] := 0.23070563;
      R_i[9,9] := 1.58302653;
      R_i[9,10] := 0.64158803;
      R_i[9,11] := -0.06970121;
      R_i[9,12] := -0.38563612;
      R_i[9,13] := -0.51418930;
      R_i[9,14] := -0.67178756;
      R_i[9,15] := 0.66275042;
      R_i[9,16] := -0.50910872;
      R_i[9,17] := 0.79785782;
      R_i[9,18] := 0.69775558;
      R_i[9,19] := -0.47073287;
      R_i[9,20] := -0.00912833;
      R_i[9,21] := 0.19374555;
      R_i[9,22] := 0.08547072;
      R_i[9,23] := -0.08412491;
      R_i[9,24] := -0.54616952;
      R_i[9,25] := 0.45187387;
      R_i[9,26] := 0.56076854;
      R_i[9,27] := 0.26952675;
      R_i[9,28] := -0.08776135;
      R_i[9,29] := 0.05690705;
      R_i[9,30] := -0.20617478;
      R_i[9,31] := -0.75883961;
      R_i[10,0] := -0.22486998;
      R_i[10,1] := 0.35497808;
      R_i[10,2] := 0.10050306;
      R_i[10,3] := 0.05792510;
      R_i[10,4] := 0.16392338;
      R_i[10,5] := -0.08192988;
      R_i[10,6] := -0.11547739;
      R_i[10,7] := -0.12439582;
      R_i[10,8] := -0.07351477;
      R_i[10,9] := 0.15080257;
      R_i[10,10] := -2.29766273;
      R_i[10,11] := 0.00198175;
      R_i[10,12] := -0.04347121;
      R_i[10,13] := 0.09138957;
      R_i[10,14] := -0.20275950;
      R_i[10,15] := 0.16711386;
      R_i[10,16] := -0.21961702;
      R_i[10,17] := 0.12318345;
      R_i[10,18] := 0.29455358;
      R_i[10,19] := 0.79191226;
      R_i[10,20] := -0.14210112;
      R_i[10,21] := -0.11408937;
      R_i[10,22] := -0.12465388;
      R_i[10,23] := -0.00793563;
      R_i[10,24] := 0.05072474;
      R_i[10,25] := -0.07968710;
      R_i[10,26] := 0.11579556;
      R_i[10,27] := -0.06528948;
      R_i[10,28] := -0.08819447;
      R_i[10,29] := -0.10903518;
      R_i[10,30] := -0.01066096;
      R_i[10,31] := -0.02178088;
      R_i[11,0] := -0.68476927;
      R_i[11,1] := 0.38765344;
      R_i[11,2] := 0.17015678;
      R_i[11,3] := -0.95622021;
      R_i[11,4] := -0.11764704;
      R_i[11,5] := 0.27207455;
      R_i[11,6] := 0.15237650;
      R_i[11,7] := -0.19831522;
      R_i[11,8] := -0.23903258;
      R_i[11,9] := 0.56660861;
      R_i[11,10] := -0.01439447;
      R_i[11,11] := -2.12028742;
      R_i[11,12] := -0.46773353;
      R_i[11,13] := 0.04793666;
      R_i[11,14] := 0.05703447;
      R_i[11,15] := 0.35312128;
      R_i[11,16] := -0.84540880;
      R_i[11,17] := 0.87920487;
      R_i[11,18] := 0.50743526;
      R_i[11,19] := 0.90020955;
      R_i[11,20] := 0.36728761;
      R_i[11,21] := -0.56907481;
      R_i[11,22] := 0.26376301;
      R_i[11,23] := -0.05402540;
      R_i[11,24] := -0.02567471;
      R_i[11,25] := -0.43724918;
      R_i[11,26] := 0.43349412;
      R_i[11,27] := -0.53790677;
      R_i[11,28] := -0.07165781;
      R_i[11,29] := 0.21291202;
      R_i[11,30] := 0.17234261;
      R_i[11,31] := -0.47796181;
      R_i[12,0] := -0.00006267;
      R_i[12,1] := 0.11495551;
      R_i[12,2] := -0.08349284;
      R_i[12,3] := -0.22248125;
      R_i[12,4] := -0.16840875;
      R_i[12,5] := 0.31274590;
      R_i[12,6] := 0.25239354;
      R_i[12,7] := -0.52599919;
      R_i[12,8] := -0.11546670;
      R_i[12,9] := 0.55316460;
      R_i[12,10] := 0.00625816;
      R_i[12,11] := -0.24307473;
      R_i[12,12] := -0.63897330;
      R_i[12,13] := 0.14157343;
      R_i[12,14] := -0.24095358;
      R_i[12,15] := -0.19407575;
      R_i[12,16] := -0.54413486;
      R_i[12,17] := -0.06198624;
      R_i[12,18] := 0.23189466;
      R_i[12,19] := 0.04720600;
      R_i[12,20] := 0.15461636;
      R_i[12,21] := 0.14028889;
      R_i[12,22] := 0.09214773;
      R_i[12,23] := -0.10140400;
      R_i[12,24] := -0.23882978;
      R_i[12,25] := -0.10693639;
      R_i[12,26] := -0.28410488;
      R_i[12,27] := 0.21555559;
      R_i[12,28] := -0.06009941;
      R_i[12,29] := 0.53120393;
      R_i[12,30] := -0.19574499;
      R_i[12,31] := 0.16197842;
      R_i[13,0] := 0.45515203;
      R_i[13,1] := -0.10936302;
      R_i[13,2] := 0.19458811;
      R_i[13,3] := -0.04792923;
      R_i[13,4] := -0.83723605;
      R_i[13,5] := -0.20762044;
      R_i[13,6] := -0.25807819;
      R_i[13,7] := -0.18988095;
      R_i[13,8] := 0.25716004;
      R_i[13,9] := 0.09518423;
      R_i[13,10] := -0.24384676;
      R_i[13,11] := 0.41867420;
      R_i[13,12] := 0.32823512;
      R_i[13,13] := 0.17112298;
      R_i[13,14] := 0.31680295;
      R_i[13,15] := 0.27173653;
      R_i[13,16] := 0.46019927;
      R_i[13,17] := -0.50040060;
      R_i[13,18] := 0.01799349;
      R_i[13,19] := -0.82000792;
      R_i[13,20] := 0.21273567;
      R_i[13,21] := -0.57424170;
      R_i[13,22] := -0.49586058;
      R_i[13,23] := 0.06957225;
      R_i[13,24] := -0.21218228;
      R_i[13,25] := 0.71526438;
      R_i[13,26] := 0.02224069;
      R_i[13,27] := 0.29907489;
      R_i[13,28] := 0.28443962;
      R_i[13,29] := 0.35106656;
      R_i[13,30] := -0.35146499;
      R_i[13,31] := 0.74115050;
      R_i[14,0] := -0.39343065;
      R_i[14,1] := 0.84045798;
      R_i[14,2] := -0.16658224;
      R_i[14,3] := -0.57521433;
      R_i[14,4] := 0.36024657;
      R_i[14,5] := -0.23194501;
      R_i[14,6] := 0.37999561;
      R_i[14,7] := -0.27919167;
      R_i[14,8] := -0.14781186;
      R_i[14,9] := 0.87664002;
      R_i[14,10] := -0.01625125;
      R_i[14,11] := -0.64787418;
      R_i[14,12] := -0.29524571;
      R_i[14,13] := -0.52903223;
      R_i[14,14] := 1.58356547;
      R_i[14,15] := 0.41859668;
      R_i[14,16] := -0.08852041;
      R_i[14,17] := 1.17931008;
      R_i[14,18] := 0.54767627;
      R_i[14,19] := -0.36519223;
      R_i[14,20] := 0.11925033;
      R_i[14,21] := 0.55935115;
      R_i[14,22] := 0.03163567;
      R_i[14,23] := -0.01081576;
      R_i[14,24] := 0.28299937;
      R_i[14,25] := -0.16483735;
      R_i[14,26] := 0.38078859;
      R_i[14,27] := -0.46654803;
      R_i[14,28] := 0.03880383;
      R_i[14,29] := -0.08690705;
      R_i[14,30] := -0.00022676;
      R_i[14,31] := -0.47718471;
      R_i[15,0] := 0.40416414;
      R_i[15,1] := -0.13255139;
      R_i[15,2] := 0.33374476;
      R_i[15,3] := -0.10753588;
      R_i[15,4] := -0.30254161;
      R_i[15,5] := -0.07972442;
      R_i[15,6] := 0.16363029;
      R_i[15,7] := 0.03312247;
      R_i[15,8] := -0.08833427;
      R_i[15,9] := 0.13303199;
      R_i[15,10] := -0.26298860;
      R_i[15,11] := -0.15168363;
      R_i[15,12] := -0.30840203;
      R_i[15,13] := -0.15638354;
      R_i[15,14] := 0.00463648;
      R_i[15,15] := -0.04008638;
      R_i[15,16] := 0.23492582;
      R_i[15,17] := 0.29362372;
      R_i[15,18] := 0.24428976;
      R_i[15,19] := -0.33830038;
      R_i[15,20] := 0.45935920;
      R_i[15,21] := -0.28399682;
      R_i[15,22] := -0.01934072;
      R_i[15,23] := -0.20523863;
      R_i[15,24] := -0.13765733;
      R_i[15,25] := -0.00695347;
      R_i[15,26] := 0.22762655;
      R_i[15,27] := -0.04855500;
      R_i[15,28] := -0.23287787;
      R_i[15,29] := 0.15384027;
      R_i[15,30] := -0.03583547;
      R_i[15,31] := -0.02649516;
      R_i[16,0] := -0.18315850;
      R_i[16,1] := 0.41206077;
      R_i[16,2] := -0.14354268;
      R_i[16,3] := -0.44737810;
      R_i[16,4] := -0.08704913;
      R_i[16,5] := 0.29804343;
      R_i[16,6] := 0.27113724;
      R_i[16,7] := -0.39558008;
      R_i[16,8] := -0.59111369;
      R_i[16,9] := 0.37798053;
      R_i[16,10] := 0.81796849;
      R_i[16,11] := -0.12820429;
      R_i[16,12] := -0.59571439;
      R_i[16,13] := -0.03124824;
      R_i[16,14] := -0.18218520;
      R_i[16,15] := 0.12198190;
      R_i[16,16] := 1.41429520;
      R_i[16,17] := 0.47617510;
      R_i[16,18] := 0.80915415;
      R_i[16,19] := 0.28500611;
      R_i[16,20] := 0.18615711;
      R_i[16,21] := 0.19952437;
      R_i[16,22] := -0.25558889;
      R_i[16,23] := -0.30694398;
      R_i[16,24] := -0.06202212;
      R_i[16,25] := 0.04830749;
      R_i[16,26] := 0.05715989;
      R_i[16,27] := -0.15100600;
      R_i[16,28] := 0.36785114;
      R_i[16,29] := 0.09471590;
      R_i[16,30] := -0.36646622;
      R_i[16,31] := 0.09723163;
      R_i[17,0] := -1.00640607;
      R_i[17,1] := 0.48862299;
      R_i[17,2] := 0.03128826;
      R_i[17,3] := 0.13596107;
      R_i[17,4] := 0.25177097;
      R_i[17,5] := 0.14061838;
      R_i[17,6] := -0.00378009;
      R_i[17,7] := 0.30384693;
      R_i[17,8] := 0.20079097;
      R_i[17,9] := 0.74782521;
      R_i[17,10] := 1.31918955;
      R_i[17,11] := -1.57991540;
      R_i[17,12] := 0.29552051;
      R_i[17,13] := -0.60454607;
      R_i[17,14] := -0.21482722;
      R_i[17,15] := 0.23917961;
      R_i[17,16] := -1.00066638;
      R_i[17,17] := 4.23797512;
      R_i[17,18] := 0.71026301;
      R_i[17,19] := 0.25954387;
      R_i[17,20] := 0.30618632;
      R_i[17,21] := -0.11564369;
      R_i[17,22] := 0.22178310;
      R_i[17,23] := -0.34120065;
      R_i[17,24] := 0.07910939;
      R_i[17,25] := -0.43872246;
      R_i[17,26] := 0.12337355;
      R_i[17,27] := -0.17299944;
      R_i[17,28] := -0.26848623;
      R_i[17,29] := -0.07663534;
      R_i[17,30] := 0.22587071;
      R_i[17,31] := -0.38025171;
      R_i[18,0] := -0.37464195;
      R_i[18,1] := 0.10491309;
      R_i[18,2] := -0.13920635;
      R_i[18,3] := -0.31322402;
      R_i[18,4] := -0.25237298;
      R_i[18,5] := 0.05783420;
      R_i[18,6] := -0.37912083;
      R_i[18,7] := -0.09298448;
      R_i[18,8] := 0.20246075;
      R_i[18,9] := 0.85220355;
      R_i[18,10] := -0.30931070;
      R_i[18,11] := -0.29023072;
      R_i[18,12] := 0.12028287;
      R_i[18,13] := -0.07692172;
      R_i[18,14] := 0.28702876;
      R_i[18,15] := 0.22447805;
      R_i[18,16] := -0.33956850;
      R_i[18,17] := 0.15055300;
      R_i[18,18] := 2.02416468;
      R_i[18,19] := 0.21693578;
      R_i[18,20] := -0.14444982;
      R_i[18,21] := 0.08650701;
      R_i[18,22] := -0.22850646;
      R_i[18,23] := 0.36052695;
      R_i[18,24] := -0.02930431;
      R_i[18,25] := 0.15847221;
      R_i[18,26] := -0.60505497;
      R_i[18,27] := 0.05648470;
      R_i[18,28] := 0.25863642;
      R_i[18,29] := -0.10821130;
      R_i[18,30] := -0.06356303;
      R_i[18,31] := 0.43008837;
      R_i[19,0] := -0.10740647;
      R_i[19,1] := -0.06138924;
      R_i[19,2] := 0.06404181;
      R_i[19,3] := 0.00516134;
      R_i[19,4] := 0.11549391;
      R_i[19,5] := 0.89629108;
      R_i[19,6] := -0.28299421;
      R_i[19,7] := -0.06409787;
      R_i[19,8] := 0.36336362;
      R_i[19,9] := 0.79763788;
      R_i[19,10] := 0.30653960;
      R_i[19,11] := -0.92557198;
      R_i[19,12] := -0.25698316;
      R_i[19,13] := -0.17551865;
      R_i[19,14] := 0.02162044;
      R_i[19,15] := 0.06503978;
      R_i[19,16] := -0.11493133;
      R_i[19,17] := 0.84433997;
      R_i[19,18] := -0.22099726;
      R_i[19,19] := -0.09091380;
      R_i[19,20] := 0.46641204;
      R_i[19,21] := -0.03867416;
      R_i[19,22] := 0.57412326;
      R_i[19,23] := -0.33754462;
      R_i[19,24] := -0.08072848;
      R_i[19,25] := 0.13773033;
      R_i[19,26] := 0.25080514;
      R_i[19,27] := -0.71225595;
      R_i[19,28] := -0.35166001;
      R_i[19,29] := -0.43134296;
      R_i[19,30] := -0.21888943;
      R_i[19,31] := 0.57688344;
      R_i[20,0] := 0.22825079;
      R_i[20,1] := 0.37793356;
      R_i[20,2] := -0.13493037;
      R_i[20,3] := -0.44883609;
      R_i[20,4] := -0.83388597;
      R_i[20,5] := 0.12293290;
      R_i[20,6] := -0.46607855;
      R_i[20,7] := -0.07845667;
      R_i[20,8] := 1.32477832;
      R_i[20,9] := 0.68255568;
      R_i[20,10] := -0.05006309;
      R_i[20,11] := -0.47491327;
      R_i[20,12] := -0.43141145;
      R_i[20,13] := 0.47282761;
      R_i[20,14] := 0.41005883;
      R_i[20,15] := -0.01599345;
      R_i[20,16] := 0.13017854;
      R_i[20,17] := 0.52654916;
      R_i[20,18] := 0.57140589;
      R_i[20,19] := 0.41956627;
      R_i[20,20] := -1.84662533;
      R_i[20,21] := -0.59662354;
      R_i[20,22] := 0.82912123;
      R_i[20,23] := -0.11413272;
      R_i[20,24] := -0.38720784;
      R_i[20,25] := -0.09421971;
      R_i[20,26] := 0.80597848;
      R_i[20,27] := 0.65747625;
      R_i[20,28] := -0.21523356;
      R_i[20,29] := 0.48304906;
      R_i[20,30] := 0.35006654;
      R_i[20,31] := -0.57040602;
      R_i[21,0] := -0.03587767;
      R_i[21,1] := 0.42292139;
      R_i[21,2] := -0.37415621;
      R_i[21,3] := -0.02178310;
      R_i[21,4] := -0.27689084;
      R_i[21,5] := 0.05678604;
      R_i[21,6] := -0.13292289;
      R_i[21,7] := 0.00694761;
      R_i[21,8] := -0.06681035;
      R_i[21,9] := 0.42398322;
      R_i[21,10] := -0.17418142;
      R_i[21,11] := -0.28406641;
      R_i[21,12] := -0.04291890;
      R_i[21,13] := 0.12964997;
      R_i[21,14] := 0.20425871;
      R_i[21,15] := 0.08085304;
      R_i[21,16] := 0.03528428;
      R_i[21,17] := 0.23000003;
      R_i[21,18] := 0.37066588;
      R_i[21,19] := -0.18582781;
      R_i[21,20] := -0.03903870;
      R_i[21,21] := 0.21170920;
      R_i[21,22] := 0.29128164;
      R_i[21,23] := -0.29781890;
      R_i[21,24] := 0.02116948;
      R_i[21,25] := -0.10276867;
      R_i[21,26] := 0.34249908;
      R_i[21,27] := 0.08698206;
      R_i[21,28] := -0.07140943;
      R_i[21,29] := -0.09261855;
      R_i[21,30] := 0.05416507;
      R_i[21,31] := -0.04114371;
      R_i[22,0] := -0.17186950;
      R_i[22,1] := 0.27311918;
      R_i[22,2] := 0.17921014;
      R_i[22,3] := -0.71519452;
      R_i[22,4] := 0.14193517;
      R_i[22,5] := -0.29420683;
      R_i[22,6] := -0.62526858;
      R_i[22,7] := -0.17676060;
      R_i[22,8] := -0.06704113;
      R_i[22,9] := 0.29654166;
      R_i[22,10] := -0.24501418;
      R_i[22,11] := 0.05814528;
      R_i[22,12] := 0.29545593;
      R_i[22,13] := -0.73224670;
      R_i[22,14] := -0.10482658;
      R_i[22,15] := 0.18565421;
      R_i[22,16] := 0.24734524;
      R_i[22,17] := 0.28190374;
      R_i[22,18] := 0.07871399;
      R_i[22,19] := 0.70523387;
      R_i[22,20] := 0.45427024;
      R_i[22,21] := -0.13728946;
      R_i[22,22] := 1.31304848;
      R_i[22,23] := -0.40054202;
      R_i[22,24] := -0.64563668;
      R_i[22,25] := -0.24695830;
      R_i[22,26] := 0.42006245;
      R_i[22,27] := -1.35477948;
      R_i[22,28] := 0.23874813;
      R_i[22,29] := -0.32546738;
      R_i[22,30] := 0.82682675;
      R_i[22,31] := 0.17273316;
      R_i[23,0] := -0.22012863;
      R_i[23,1] := 0.04423183;
      R_i[23,2] := 0.83607686;
      R_i[23,3] := -0.10190780;
      R_i[23,4] := -0.44084197;
      R_i[23,5] := -0.01347674;
      R_i[23,6] := -0.39046064;
      R_i[23,7] := -0.45612475;
      R_i[23,8] := -0.52376109;
      R_i[23,9] := 0.23790218;
      R_i[23,10] := -0.20900583;
      R_i[23,11] := -0.55885947;
      R_i[23,12] := -0.08895622;
      R_i[23,13] := 0.25092366;
      R_i[23,14] := 0.34155697;
      R_i[23,15] := 0.34225461;
      R_i[23,16] := 0.37864837;
      R_i[23,17] := 0.06985009;
      R_i[23,18] := 0.25320885;
      R_i[23,19] := -0.71266365;
      R_i[23,20] := -0.08440322;
      R_i[23,21] := -0.22635168;
      R_i[23,22] := -0.09268820;
      R_i[23,23] := 0.76479942;
      R_i[23,24] := 0.17106181;
      R_i[23,25] := -0.39618358;
      R_i[23,26] := 1.07378483;
      R_i[23,27] := -0.60030353;
      R_i[23,28] := 0.43353710;
      R_i[23,29] := 0.37375939;
      R_i[23,30] := 0.31260803;
      R_i[23,31] := 0.36026886;
      R_i[24,0] := 0.43552378;
      R_i[24,1] := -0.60323244;
      R_i[24,2] := -0.22056930;
      R_i[24,3] := 0.30780360;
      R_i[24,4] := -0.41191232;
      R_i[24,5] := -0.07733422;
      R_i[24,6] := -0.47244716;
      R_i[24,7] := 0.21977623;
      R_i[24,8] := 0.28462246;
      R_i[24,9] := 0.17637153;
      R_i[24,10] := -0.32458791;
      R_i[24,11] := 0.43863761;
      R_i[24,12] := 0.33493611;
      R_i[24,13] := 0.35019112;
      R_i[24,14] := 0.32484850;
      R_i[24,15] := -0.09011348;
      R_i[24,16] := 0.55679053;
      R_i[24,17] := -0.32762069;
      R_i[24,18] := -0.21257828;
      R_i[24,19] := -0.55349809;
      R_i[24,20] := -0.09330451;
      R_i[24,21] := 0.01841493;
      R_i[24,22] := 0.18566658;
      R_i[24,23] := -0.02519841;
      R_i[24,24] := 0.10400505;
      R_i[24,25] := 0.38245302;
      R_i[24,26] := 0.64739758;
      R_i[24,27] := 0.04741986;
      R_i[24,28] := 0.16349974;
      R_i[24,29] := 0.07289705;
      R_i[24,30] := -0.09029396;
      R_i[24,31] := -0.02031578;
      R_i[25,0] := -0.53194910;
      R_i[25,1] := 0.02412759;
      R_i[25,2] := -1.21617222;
      R_i[25,3] := -0.65800297;
      R_i[25,4] := -0.57248634;
      R_i[25,5] := -1.31935811;
      R_i[25,6] := 1.16315258;
      R_i[25,7] := 0.61346394;
      R_i[25,8] := 0.76240295;
      R_i[25,9] := -0.15611924;
      R_i[25,10] := 0.95619309;
      R_i[25,11] := 0.68118155;
      R_i[25,12] := 0.13858624;
      R_i[25,13] := -0.34527764;
      R_i[25,14] := -0.45235732;
      R_i[25,15] := 0.29673636;
      R_i[25,16] := 0.34407869;
      R_i[25,17] := -0.34264007;
      R_i[25,18] := 0.01217187;
      R_i[25,19] := -0.33046424;
      R_i[25,20] := 0.09931978;
      R_i[25,21] := -1.01859987;
      R_i[25,22] := 0.89789706;
      R_i[25,23] := 0.02949729;
      R_i[25,24] := -0.00726639;
      R_i[25,25] := -0.58121955;
      R_i[25,26] := -0.61388236;
      R_i[25,27] := -0.29241377;
      R_i[25,28] := 0.46526292;
      R_i[25,29] := -0.07431906;
      R_i[25,30] := -0.26869741;
      R_i[25,31] := -0.67653674;
      R_i[26,0] := -0.34057721;
      R_i[26,1] := -0.09010746;
      R_i[26,2] := -0.31317073;
      R_i[26,3] := -0.97618186;
      R_i[26,4] := 0.82685155;
      R_i[26,5] := -4.58021116;
      R_i[26,6] := 1.36010897;
      R_i[26,7] := -0.47619432;
      R_i[26,8] := 2.03470421;
      R_i[26,9] := -0.53427881;
      R_i[26,10] := -0.13629383;
      R_i[26,11] := -0.13242298;
      R_i[26,12] := 0.28095043;
      R_i[26,13] := 0.95876056;
      R_i[26,14] := 0.48941121;
      R_i[26,15] := 0.19460116;
      R_i[26,16] := 0.16457404;
      R_i[26,17] := -0.65959787;
      R_i[26,18] := 0.06110868;
      R_i[26,19] := 1.14294267;
      R_i[26,20] := -0.10814787;
      R_i[26,21] := 0.74087745;
      R_i[26,22] := -2.00501585;
      R_i[26,23] := 0.24415712;
      R_i[26,24] := -3.70227790;
      R_i[26,25] := -1.56724083;
      R_i[26,26] := -3.67185569;
      R_i[26,27] := 1.17687500;
      R_i[26,28] := -1.88574040;
      R_i[26,29] := 0.23438171;
      R_i[26,30] := 0.92084801;
      R_i[26,31] := 1.74960470;
      R_i[27,0] := 0.08044783;
      R_i[27,1] := -0.04984543;
      R_i[27,2] := -0.24893922;
      R_i[27,3] := -0.21227036;
      R_i[27,4] := -0.15274289;
      R_i[27,5] := 0.01640888;
      R_i[27,6] := -0.53605032;
      R_i[27,7] := 0.24002981;
      R_i[27,8] := 0.20014673;
      R_i[27,9] := -0.02934171;
      R_i[27,10] := -0.08759493;
      R_i[27,11] := 0.63402885;
      R_i[27,12] := 0.01651026;
      R_i[27,13] := 0.09693064;
      R_i[27,14] := 0.29044932;
      R_i[27,15] := -0.28162980;
      R_i[27,16] := 0.29138079;
      R_i[27,17] := -0.08596911;
      R_i[27,18] := 0.06656250;
      R_i[27,19] := -0.42018428;
      R_i[27,20] := -0.07639185;
      R_i[27,21] := 0.54837906;
      R_i[27,22] := 0.00699990;
      R_i[27,23] := 0.57944459;
      R_i[27,24] := -0.32708910;
      R_i[27,25] := -0.05541108;
      R_i[27,26] := 0.04765628;
      R_i[27,27] := -0.35345450;
      R_i[27,28] := -0.00601142;
      R_i[27,29] := 0.29992521;
      R_i[27,30] := -0.31607386;
      R_i[27,31] := 0.41685253;
      R_i[28,0] := -0.49491948;
      R_i[28,1] := 0.69275510;
      R_i[28,2] := -0.44414425;
      R_i[28,3] := 0.08284695;
      R_i[28,4] := 0.19715372;
      R_i[28,5] := -0.11869717;
      R_i[28,6] := 0.43726832;
      R_i[28,7] := 0.06932707;
      R_i[28,8] := 0.62274700;
      R_i[28,9] := 0.61477602;
      R_i[28,10] := -0.22220217;
      R_i[28,11] := -0.68593425;
      R_i[28,12] := 0.23542540;
      R_i[28,13] := -0.48637852;
      R_i[28,14] := -0.01314360;
      R_i[28,15] := -0.17047518;
      R_i[28,16] := -0.11696369;
      R_i[28,17] := -0.07707114;
      R_i[28,18] := -0.53148073;
      R_i[28,19] := -0.48331252;
      R_i[28,20] := 0.27698728;
      R_i[28,21] := 0.10087790;
      R_i[28,22] := 0.19291788;
      R_i[28,23] := 0.12205473;
      R_i[28,24] := 0.53354186;
      R_i[28,25] := -0.27771723;
      R_i[28,26] := 0.42416579;
      R_i[28,27] := -0.06338947;
      R_i[28,28] := 0.98868507;
      R_i[28,29] := -0.42105702;
      R_i[28,30] := 0.47273302;
      R_i[28,31] := -0.45523530;
      R_i[29,0] := -0.13489522;
      R_i[29,1] := 0.51308405;
      R_i[29,2] := -0.49689013;
      R_i[29,3] := 0.31196389;
      R_i[29,4] := 0.09658425;
      R_i[29,5] := -0.15041424;
      R_i[29,6] := -0.12860303;
      R_i[29,7] := -0.41769654;
      R_i[29,8] := -0.05634471;
      R_i[29,9] := 0.52302653;
      R_i[29,10] := -0.15310770;
      R_i[29,11] := -0.08379830;
      R_i[29,12] := -0.71298873;
      R_i[29,13] := 0.46460947;
      R_i[29,14] := -0.50818044;
      R_i[29,15] := -0.18320751;
      R_i[29,16] := -0.18891114;
      R_i[29,17] := -0.08116098;
      R_i[29,18] := -0.15882139;
      R_i[29,19] := 0.49746534;
      R_i[29,20] := -0.00006439;
      R_i[29,21] := -0.17106183;
      R_i[29,22] := 0.39743838;
      R_i[29,23] := -0.54420906;
      R_i[29,24] := -0.16971061;
      R_i[29,25] := -0.09644472;
      R_i[29,26] := -0.08555771;
      R_i[29,27] := 0.61670017;
      R_i[29,28] := -0.41806170;
      R_i[29,29] := -1.22626007;
      R_i[29,30] := 0.23427823;
      R_i[29,31] := -0.08933322;
      R_i[30,0] := 0.23229377;
      R_i[30,1] := -0.09377514;
      R_i[30,2] := -0.15244894;
      R_i[30,3] := -0.28959605;
      R_i[30,4] := -0.06356224;
      R_i[30,5] := 1.10057747;
      R_i[30,6] := 1.41015232;
      R_i[30,7] := -0.03006789;
      R_i[30,8] := 0.83613080;
      R_i[30,9] := 0.40837902;
      R_i[30,10] := 0.29028663;
      R_i[30,11] := -0.57439047;
      R_i[30,12] := 0.13172196;
      R_i[30,13] := -0.65824729;
      R_i[30,14] := -0.16851293;
      R_i[30,15] := 0.90380752;
      R_i[30,16] := 0.52042270;
      R_i[30,17] := 0.29417369;
      R_i[30,18] := -0.55374843;
      R_i[30,19] := -0.35138455;
      R_i[30,20] := 0.65716529;
      R_i[30,21] := 0.20918609;
      R_i[30,22] := -0.37513319;
      R_i[30,23] := 0.34159601;
      R_i[30,24] := 0.76639676;
      R_i[30,25] := 0.04368726;
      R_i[30,26] := 1.03825164;
      R_i[30,27] := -0.33677122;
      R_i[30,28] := 0.17882183;
      R_i[30,29] := -0.34231511;
      R_i[30,30] := -1.53495800;
      R_i[30,31] := -0.26110783;
      R_i[31,0] := 0.07627262;
      R_i[31,1] := -0.09820248;
      R_i[31,2] := 0.34046781;
      R_i[31,3] := 0.15434141;
      R_i[31,4] := -0.39283854;
      R_i[31,5] := -0.53014910;
      R_i[31,6] := 0.12517647;
      R_i[31,7] := -0.19974521;
      R_i[31,8] := -0.38137439;
      R_i[31,9] := 0.06925905;
      R_i[31,10] := -0.10800895;
      R_i[31,11] := -0.15322471;
      R_i[31,12] := 0.01474523;
      R_i[31,13] := -0.29487473;
      R_i[31,14] := -0.12196346;
      R_i[31,15] := 0.32134181;
      R_i[31,16] := 0.65321797;
      R_i[31,17] := 0.51920581;
      R_i[31,18] := -0.22277474;
      R_i[31,19] := -0.89724433;
      R_i[31,20] := 0.93045974;
      R_i[31,21] := -0.47842970;
      R_i[31,22] := 0.07066959;
      R_i[31,23] := 0.17044164;
      R_i[31,24] := -0.76020449;
      R_i[31,25] := -0.17217229;
      R_i[31,26] := 0.29752541;
      R_i[31,27] := -0.23179249;
      R_i[31,28] := 0.18026105;
      R_i[31,29] := -0.03253032;
      R_i[31,30] := 0.36841980;
      R_i[31,31] := 0.94482881;
      R_f[0,0] := 0.14747813;
      R_f[0,1] := -0.22737564;
      R_f[0,2] := -0.55617356;
      R_f[0,3] := -0.29175285;
      R_f[0,4] := 1.86681211;
      R_f[0,5] := -0.66840529;
      R_f[0,6] := -0.30587864;
      R_f[0,7] := 0.32244295;
      R_f[0,8] := 0.47369158;
      R_f[0,9] := -0.76385182;
      R_f[0,10] := -0.43740147;
      R_f[0,11] := -0.34984481;
      R_f[0,12] := 0.32688046;
      R_f[0,13] := -0.95900995;
      R_f[0,14] := 1.00176489;
      R_f[0,15] := -0.45252505;
      R_f[0,16] := -0.60881567;
      R_f[0,17] := -0.21773516;
      R_f[0,18] := -0.78758121;
      R_f[0,19] := -0.20532016;
      R_f[0,20] := -0.41188270;
      R_f[0,21] := -0.13742571;
      R_f[0,22] := -0.98679680;
      R_f[0,23] := -0.91927212;
      R_f[0,24] := 0.74508965;
      R_f[0,25] := 1.80925202;
      R_f[0,26] := -0.02046647;
      R_f[0,27] := 1.65381408;
      R_f[0,28] := -1.33271313;
      R_f[0,29] := -0.06231561;
      R_f[0,30] := 1.22926712;
      R_f[0,31] := 0.65283728;
      R_f[1,0] := -0.02189952;
      R_f[1,1] := 0.97953767;
      R_f[1,2] := 0.11793982;
      R_f[1,3] := -0.67327839;
      R_f[1,4] := 0.47492605;
      R_f[1,5] := 0.39999291;
      R_f[1,6] := -0.10774019;
      R_f[1,7] := 0.00958368;
      R_f[1,8] := -0.38735765;
      R_f[1,9] := -0.79148316;
      R_f[1,10] := 0.06264576;
      R_f[1,11] := -0.03151221;
      R_f[1,12] := -0.21603286;
      R_f[1,13] := -0.32396203;
      R_f[1,14] := 0.54240441;
      R_f[1,15] := 0.16125287;
      R_f[1,16] := -0.21920511;
      R_f[1,17] := -0.13962117;
      R_f[1,18] := 0.12546167;
      R_f[1,19] := 0.12239122;
      R_f[1,20] := -0.41273832;
      R_f[1,21] := -0.30105165;
      R_f[1,22] := 0.04989962;
      R_f[1,23] := 0.13209695;
      R_f[1,24] := 0.44726422;
      R_f[1,25] := 0.26851365;
      R_f[1,26] := 0.01210188;
      R_f[1,27] := 0.10423112;
      R_f[1,28] := -0.29235309;
      R_f[1,29] := 0.39567059;
      R_f[1,30] := 0.72519821;
      R_f[1,31] := 0.39522207;
      R_f[2,0] := 0.17898594;
      R_f[2,1] := -0.60384291;
      R_f[2,2] := -0.47823650;
      R_f[2,3] := -0.30635026;
      R_f[2,4] := 0.74705386;
      R_f[2,5] := -0.70426100;
      R_f[2,6] := 0.58224726;
      R_f[2,7] := 0.01940207;
      R_f[2,8] := -0.15389726;
      R_f[2,9] := -0.58458942;
      R_f[2,10] := 0.13777883;
      R_f[2,11] := -0.14377870;
      R_f[2,12] := -0.28986457;
      R_f[2,13] := -1.08470559;
      R_f[2,14] := -0.19216579;
      R_f[2,15] := -0.37692460;
      R_f[2,16] := 0.05644243;
      R_f[2,17] := 0.46512228;
      R_f[2,18] := -0.92777926;
      R_f[2,19] := -0.54135638;
      R_f[2,20] := 0.06985910;
      R_f[2,21] := -0.14253607;
      R_f[2,22] := -0.14822762;
      R_f[2,23] := 0.09599750;
      R_f[2,24] := 0.61374724;
      R_f[2,25] := 0.71291065;
      R_f[2,26] := 0.61632323;
      R_f[2,27] := 3.54531908;
      R_f[2,28] := -0.24208929;
      R_f[2,29] := 0.01456270;
      R_f[2,30] := 1.36325657;
      R_f[2,31] := 0.63486433;
      R_f[3,0] := 0.39719501;
      R_f[3,1] := 0.84666193;
      R_f[3,2] := -0.32044360;
      R_f[3,3] := 0.82361579;
